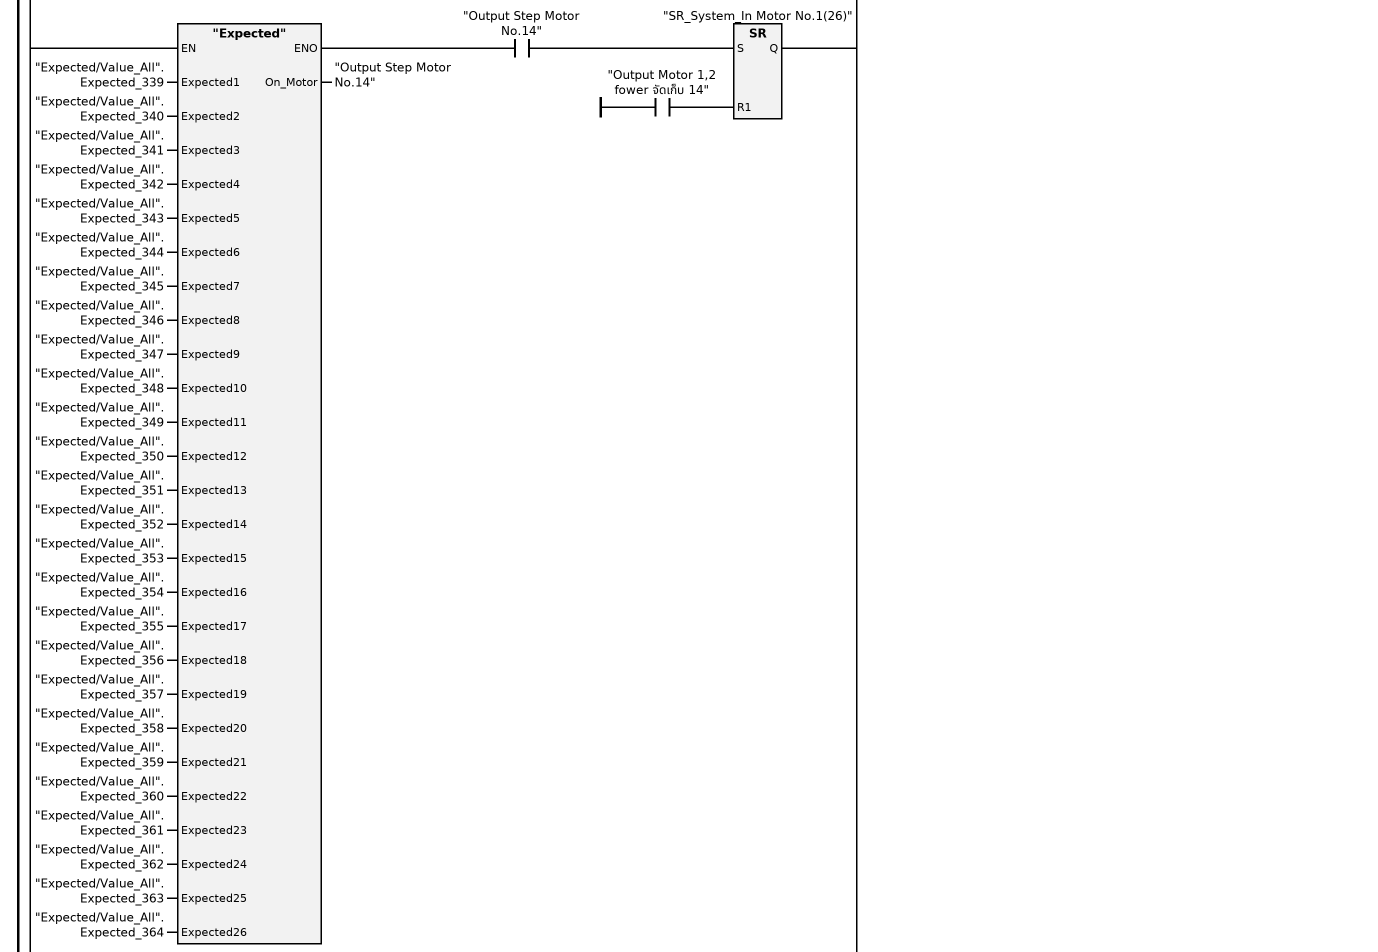
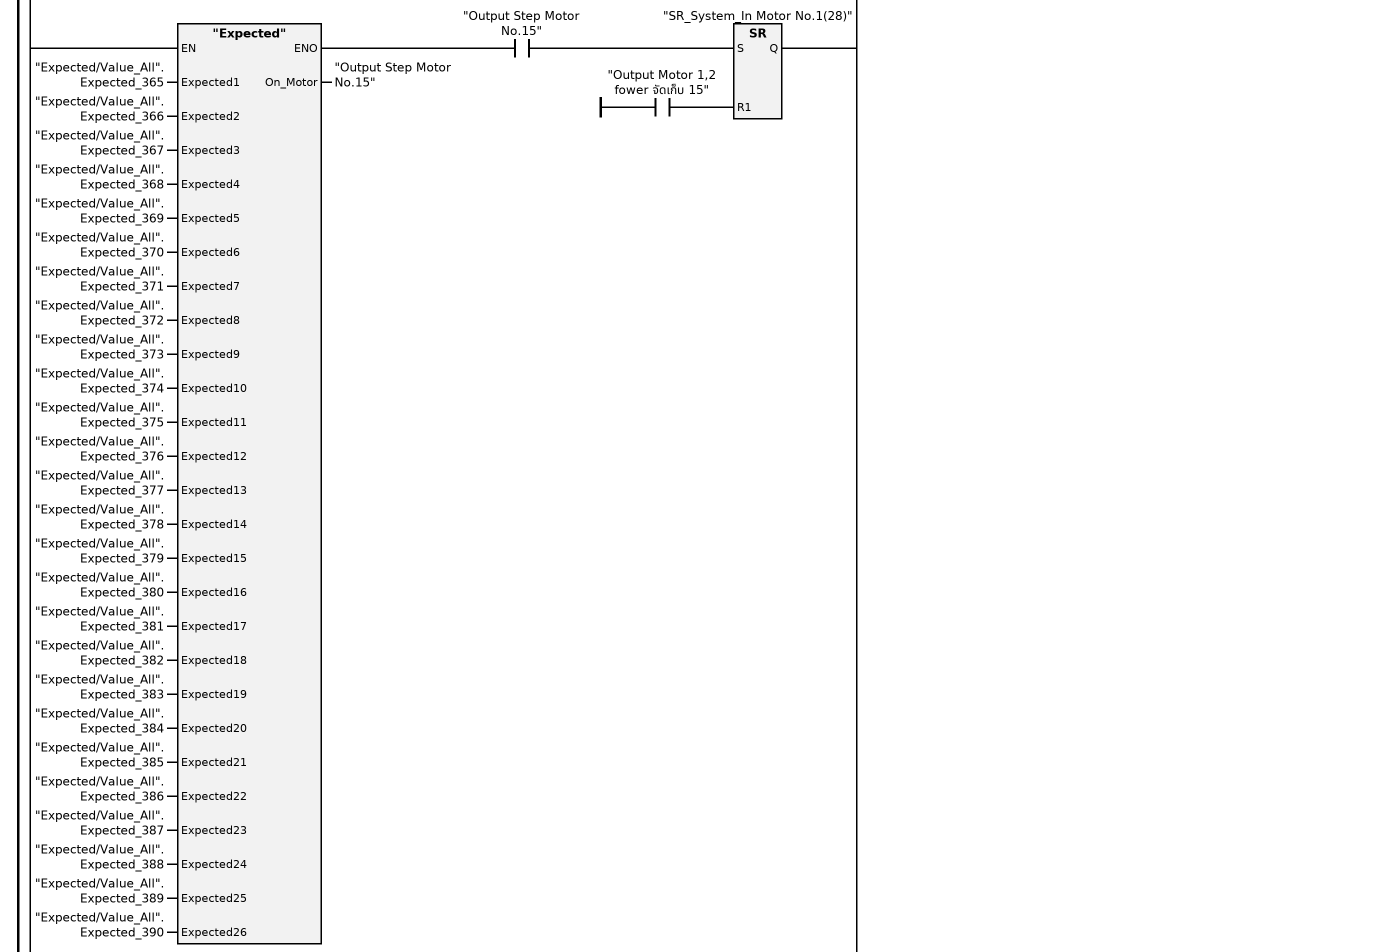
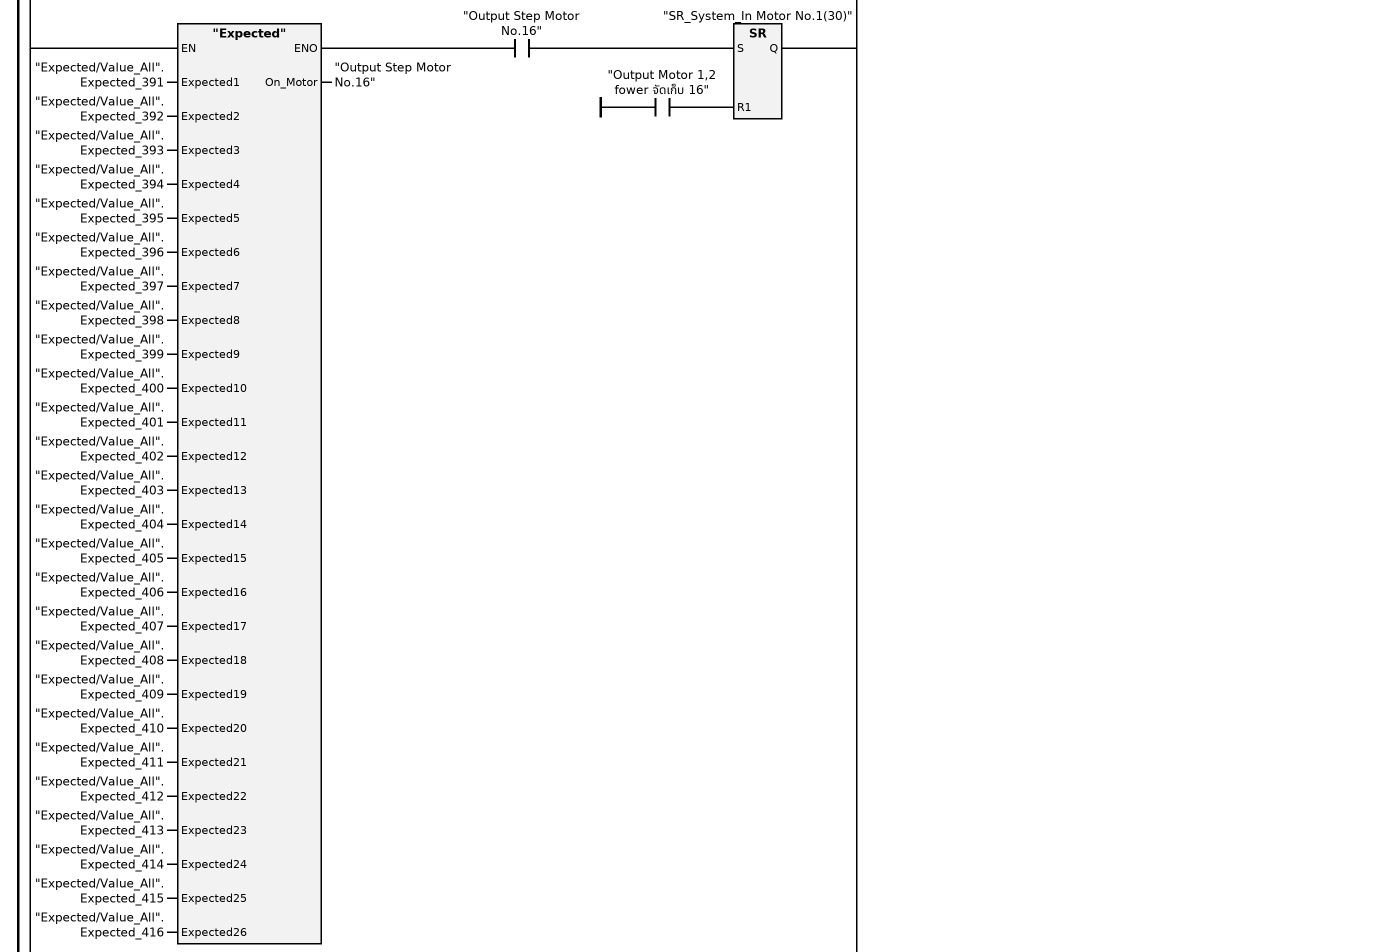
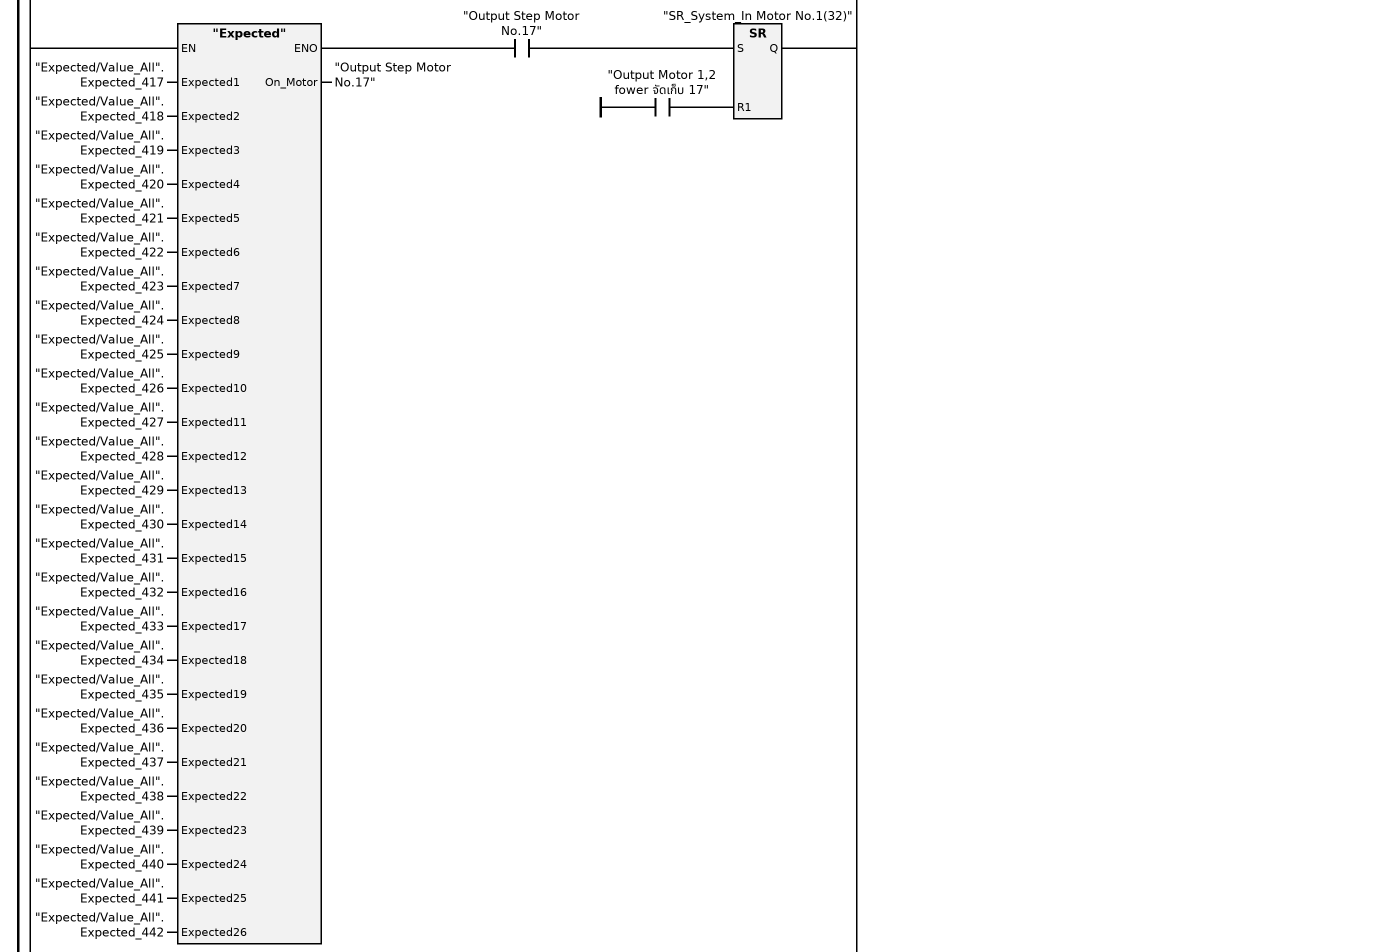
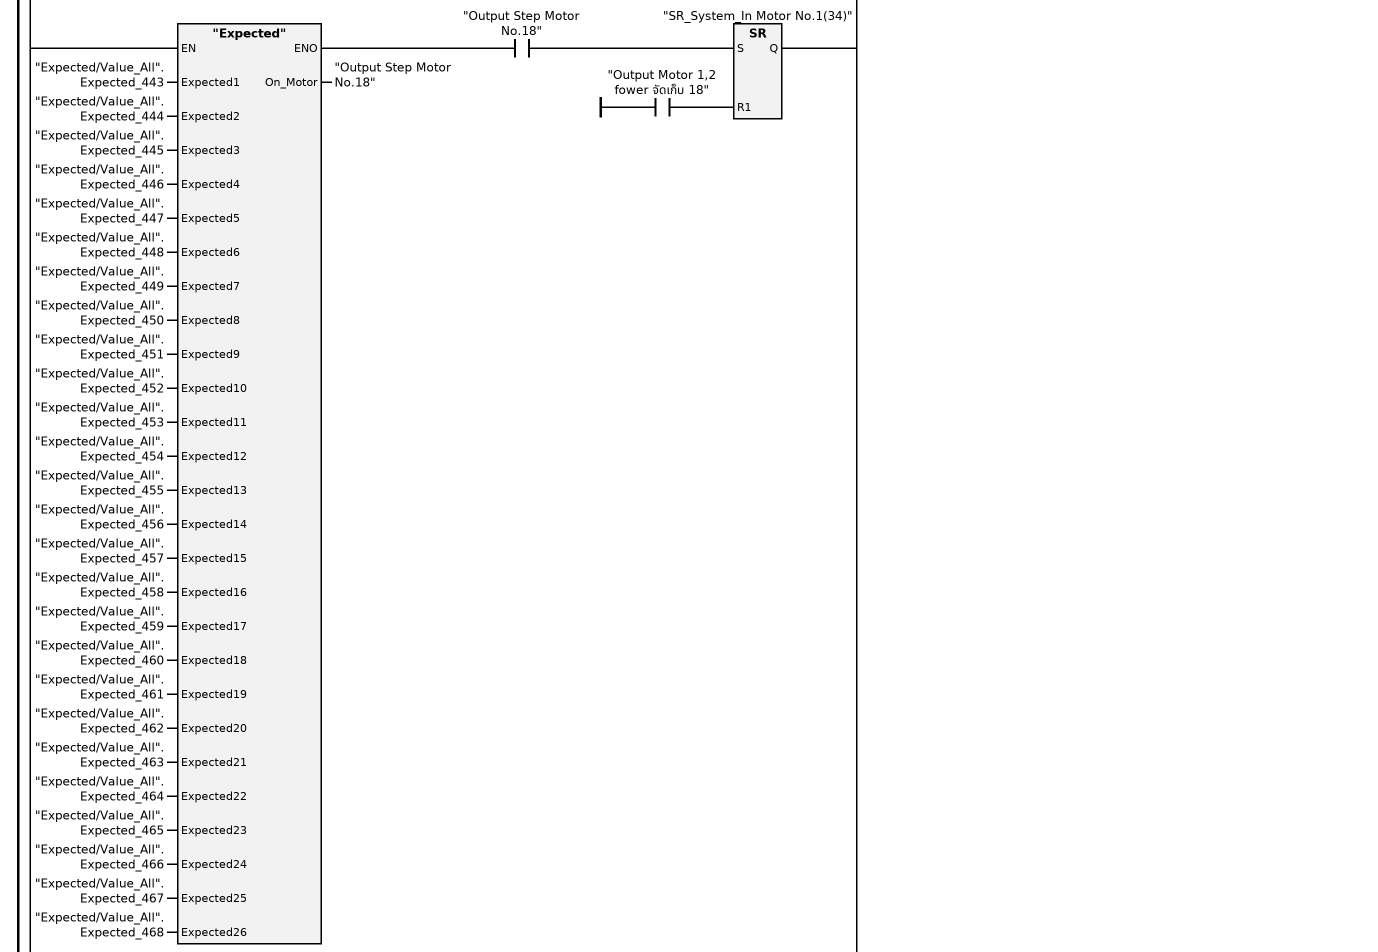
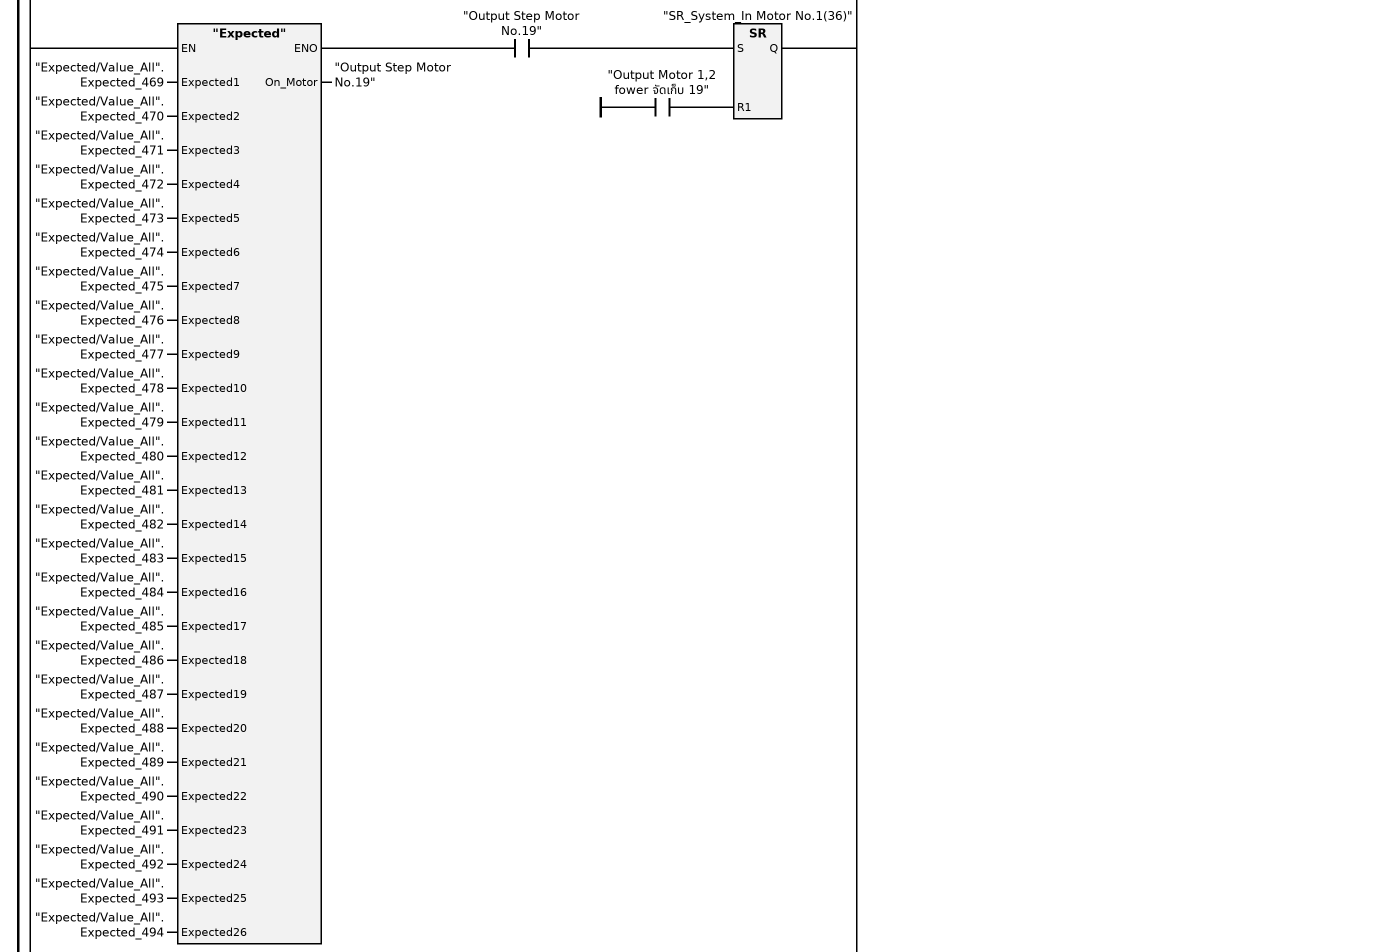
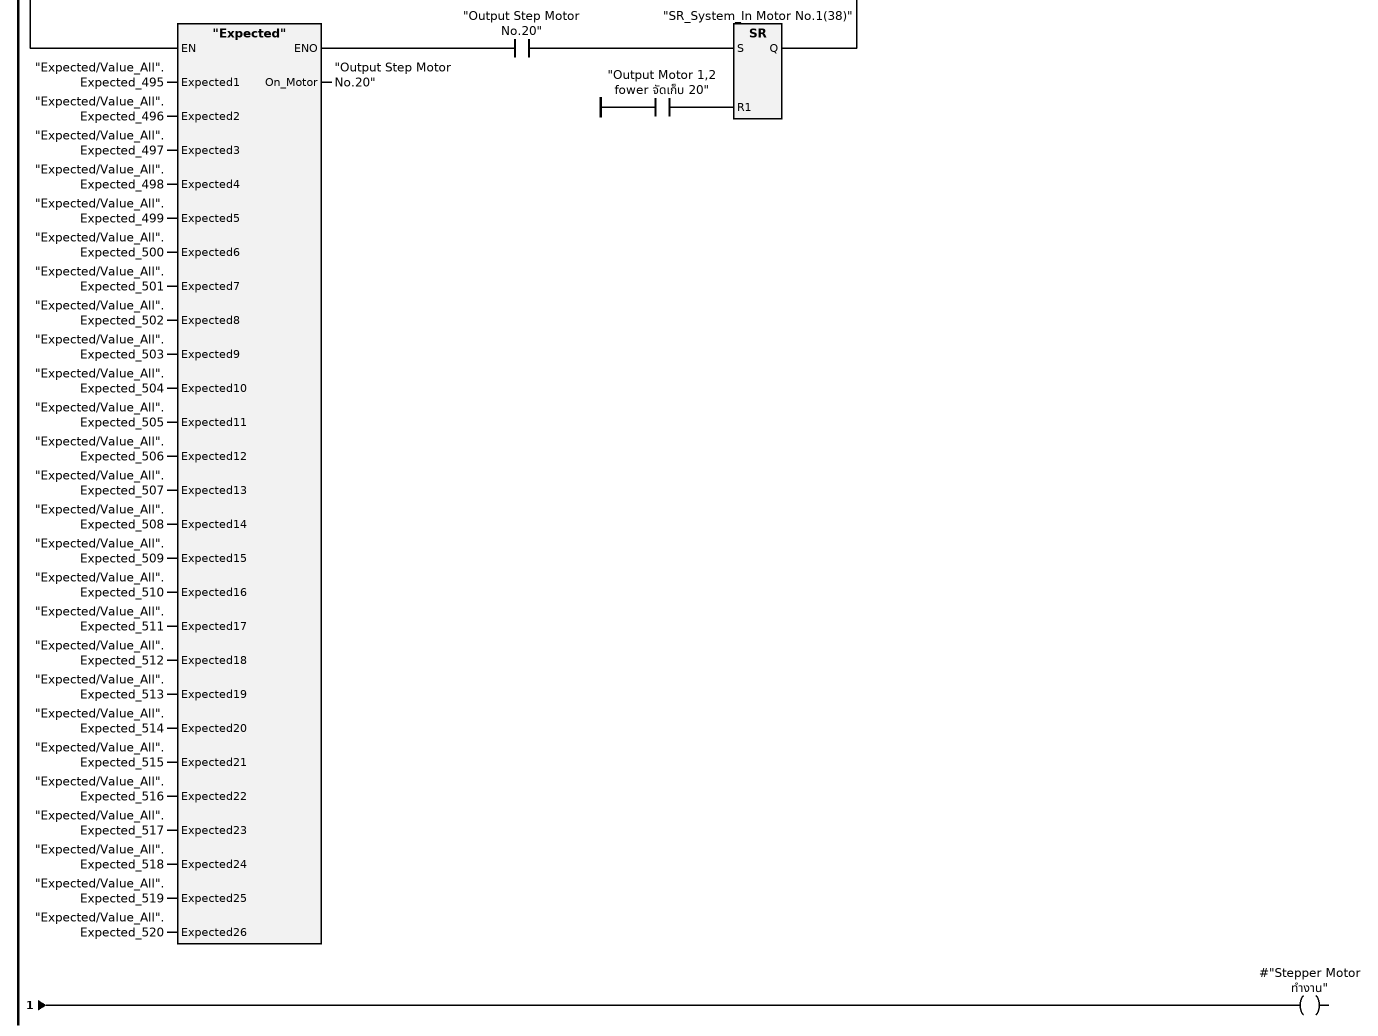
   RUNG wire#powerrail
      "Expected"(Expected1 := "Expected/Value_All".Expected_1, Expected2 := "Expected/Value_All".Expected_2, Expected3 := "Expected/Value_All".Expected_3, Expected4 := "Expected/Value_All".Expected_4, Expected5 := "Expected/Value_All".Expected_5, Expected6 := "Expected/Value_All".Expected_6, Expected7 := "Expected/Value_All".Expected_7, Expected8 := "Expected/Value_All".Expected_8, Expected9 := "Expected/Value_All".Expected_9, Expected10 := "Expected/Value_All".Expected_10, Expected11 := "Expected/Value_All".Expected_11, Expected12 := "Expected/Value_All".Expected_12, Expected13 := "Expected/Value_All".Expected_13, Expected14 := "Expected/Value_All".Expected_14, Expected15 := "Expected/Value_All".Expected_15, Expected16 := "Expected/Value_All".Expected_16, Expected17 := "Expected/Value_All".Expected_17, Expected18 := "Expected/Value_All".Expected_18, Expected19 := "Expected/Value_All".Expected_19, Expected20 := "Expected/Value_All".Expected_20, Expected21 := "Expected/Value_All".Expected_21, Expected22 := "Expected/Value_All".Expected_22, Expected23 := "Expected/Value_All".Expected_23, Expected24 := "Expected/Value_All".Expected_24, Expected25 := "Expected/Value_All".Expected_25, Expected26 := "Expected/Value_All".Expected_26, On_Motor => "Output Step Motor No.1")
      Contact( "Output Step Motor No.1" )
      S_SR(operand := "SR_System_In Motor No.1", r1 := wire#w1)
      wire#w2
      "test หลังเคลื่อนที่มาตำแหน่งปล่อยกล่องยา"()
      Contact( "หมุนไปตำแหต่งปล่อยกล่องยา" )
      Coil( #"Stepper Motor  ทำงาน" )
   END_RUNG
   RUNG wire#powerrail
      Contact( "Output Motor 1,2 fower จัดเก็บ 1" )
   END_RUNG wire#w1
   RUNG wire#powerrail
      "Expected"(Expected1 := "Expected/Value_All".Expected_27, Expected2 := "Expected/Value_All".Expected_28, Expected3 := "Expected/Value_All".Expected_29, Expected4 := "Expected/Value_All".Expected_30, Expected5 := "Expected/Value_All".Expected_31, Expected6 := "Expected/Value_All".Expected_32, Expected7 := "Expected/Value_All".Expected_33, Expected8 := "Expected/Value_All".Expected_34, Expected9 := "Expected/Value_All".Expected_35, Expected10 := "Expected/Value_All".Expected_36, Expected11 := "Expected/Value_All".Expected_37, Expected12 := "Expected/Value_All".Expected_38, Expected13 := "Expected/Value_All".Expected_39, Expected14 := "Expected/Value_All".Expected_40, Expected15 := "Expected/Value_All".Expected_41, Expected16 := "Expected/Value_All".Expected_42, Expected17 := "Expected/Value_All".Expected_43, Expected18 := "Expected/Value_All".Expected_44, Expected19 := "Expected/Value_All".Expected_45, Expected20 := "Expected/Value_All".Expected_46, Expected21 := "Expected/Value_All".Expected_47, Expected22 := "Expected/Value_All".Expected_48, Expected23 := "Expected/Value_All".Expected_49, Expected24 := "Expected/Value_All".Expected_50, Expected25 := "Expected/Value_All".Expected_51, Expected26 := "Expected/Value_All".Expected_52, On_Motor => "Output Step Motor No.2")
      Contact( "Output Step Motor No.2" )
      S_SR(operand := "SR_System_In Motor No.1(2)", r1 := wire#w3)
   END_RUNG wire#w2
   RUNG wire#powerrail
      Contact( "Output Motor 1,2 fower จัดเก็บ 2" )
   END_RUNG wire#w3
   RUNG wire#powerrail
      "Expected"(Expected1 := "Expected/Value_All".Expected_53, Expected2 := "Expected/Value_All".Expected_54, Expected3 := "Expected/Value_All".Expected_55, Expected4 := "Expected/Value_All".Expected_56, Expected5 := "Expected/Value_All".Expected_57, Expected6 := "Expected/Value_All".Expected_58, Expected7 := "Expected/Value_All".Expected_59, Expected8 := "Expected/Value_All".Expected_60, Expected9 := "Expected/Value_All".Expected_61, Expected10 := "Expected/Value_All".Expected_62, Expected11 := "Expected/Value_All".Expected_63, Expected12 := "Expected/Value_All".Expected_64, Expected13 := "Expected/Value_All".Expected_65, Expected14 := "Expected/Value_All".Expected_66, Expected15 := "Expected/Value_All".Expected_67, Expected16 := "Expected/Value_All".Expected_68, Expected17 := "Expected/Value_All".Expected_69, Expected18 := "Expected/Value_All".Expected_70, Expected19 := "Expected/Value_All".Expected_71, Expected20 := "Expected/Value_All".Expected_72, Expected21 := "Expected/Value_All".Expected_73, Expected22 := "Expected/Value_All".Expected_74, Expected23 := "Expected/Value_All".Expected_75, Expected24 := "Expected/Value_All".Expected_76, Expected25 := "Expected/Value_All".Expected_77, Expected26 := "Expected/Value_All".Expected_78, On_Motor => "Output Step Motor No.3")
      Contact( "Output Step Motor No.3" )
      S_SR(operand := "SR_System_In Motor No.1(4)", r1 := wire#w4)
   END_RUNG wire#w2
   RUNG wire#powerrail
      Contact( "Output Motor 1,2 fower จัดเก็บ 3" )
   END_RUNG wire#w4
   RUNG wire#powerrail
      "Expected"(Expected1 := "Expected/Value_All".Expected_79, Expected2 := "Expected/Value_All".Expected_80, Expected3 := "Expected/Value_All".Expected_81, Expected4 := "Expected/Value_All".Expected_82, Expected5 := "Expected/Value_All".Expected_83, Expected6 := "Expected/Value_All".Expected_84, Expected7 := "Expected/Value_All".Expected_85, Expected8 := "Expected/Value_All".Expected_86, Expected9 := "Expected/Value_All".Expected_87, Expected10 := "Expected/Value_All".Expected_88, Expected11 := "Expected/Value_All".Expected_89, Expected12 := "Expected/Value_All".Expected_90, Expected13 := "Expected/Value_All".Expected_91, Expected14 := "Expected/Value_All".Expected_92, Expected15 := "Expected/Value_All".Expected_93, Expected16 := "Expected/Value_All".Expected_94, Expected17 := "Expected/Value_All".Expected_95, Expected18 := "Expected/Value_All".Expected_96, Expected19 := "Expected/Value_All".Expected_97, Expected20 := "Expected/Value_All".Expected_98, Expected21 := "Expected/Value_All".Expected_99, Expected22 := "Expected/Value_All".Expected_100, Expected23 := "Expected/Value_All".Expected_101, Expected24 := "Expected/Value_All".Expected_102, Expected25 := "Expected/Value_All".Expected_103, Expected26 := "Expected/Value_All".Expected_104, On_Motor => "Output Step Motor No.4")
      Contact( "Output Step Motor No.4" )
      S_SR(operand := "SR_System_In Motor No.1(6)", r1 := wire#w5)
   END_RUNG wire#w2
   RUNG wire#powerrail
      Contact( "Output Motor 1,2 fower จัดเก็บ 4" )
   END_RUNG wire#w5
   RUNG wire#powerrail
      "Expected"(Expected1 := "Expected/Value_All".Expected_105, Expected2 := "Expected/Value_All".Expected_106, Expected3 := "Expected/Value_All".Expected_107, Expected4 := "Expected/Value_All".Expected_108, Expected5 := "Expected/Value_All".Expected_109, Expected6 := "Expected/Value_All".Expected_110, Expected7 := "Expected/Value_All".Expected_111, Expected8 := "Expected/Value_All".Expected_112, Expected9 := "Expected/Value_All".Expected_113, Expected10 := "Expected/Value_All".Expected_114, Expected11 := "Expected/Value_All".Expected_115, Expected12 := "Expected/Value_All".Expected_116, Expected13 := "Expected/Value_All".Expected_117, Expected14 := "Expected/Value_All".Expected_118, Expected15 := "Expected/Value_All".Expected_119, Expected16 := "Expected/Value_All".Expected_120, Expected17 := "Expected/Value_All".Expected_121, Expected18 := "Expected/Value_All".Expected_122, Expected19 := "Expected/Value_All".Expected_123, Expected20 := "Expected/Value_All".Expected_124, Expected21 := "Expected/Value_All".Expected_125, Expected22 := "Expected/Value_All".Expected_126, Expected23 := "Expected/Value_All".Expected_127, Expected24 := "Expected/Value_All".Expected_128, Expected25 := "Expected/Value_All".Expected_129, Expected26 := "Expected/Value_All".Expected_130, On_Motor => "Output Step Motor No.5")
      Contact( "Output Step Motor No.5" )
      S_SR(operand := "SR_System_In Motor No.1(8)", r1 := wire#w6)
   END_RUNG wire#w2
   RUNG wire#powerrail
      Contact( "Output Motor 1,2 fower จัดเก็บ 5" )
   END_RUNG wire#w6
   RUNG wire#powerrail
      "Expected"(Expected1 := "Expected/Value_All".Expected_131, Expected2 := "Expected/Value_All".Expected_132, Expected3 := "Expected/Value_All".Expected_133, Expected4 := "Expected/Value_All".Expected_134, Expected5 := "Expected/Value_All".Expected_135, Expected6 := "Expected/Value_All".Expected_136, Expected7 := "Expected/Value_All".Expected_137, Expected8 := "Expected/Value_All".Expected_138, Expected9 := "Expected/Value_All".Expected_139, Expected10 := "Expected/Value_All".Expected_140, Expected11 := "Expected/Value_All".Expected_141, Expected12 := "Expected/Value_All".Expected_142, Expected13 := "Expected/Value_All".Expected_143, Expected14 := "Expected/Value_All".Expected_144, Expected15 := "Expected/Value_All".Expected_145, Expected16 := "Expected/Value_All".Expected_146, Expected17 := "Expected/Value_All".Expected_147, Expected18 := "Expected/Value_All".Expected_148, Expected19 := "Expected/Value_All".Expected_149, Expected20 := "Expected/Value_All".Expected_150, Expected21 := "Expected/Value_All".Expected_151, Expected22 := "Expected/Value_All".Expected_152, Expected23 := "Expected/Value_All".Expected_153, Expected24 := "Expected/Value_All".Expected_154, Expected25 := "Expected/Value_All".Expected_155, Expected26 := "Expected/Value_All".Expected_156, On_Motor => "Output Step Motor No.6")
      Contact( "Output Step Motor No.6" )
      S_SR(operand := "SR_System_In Motor No.1(10)", r1 := wire#w7)
   END_RUNG wire#w2
   RUNG wire#powerrail
      Contact( "Output Motor 1,2 fower จัดเก็บ 6" )
   END_RUNG wire#w7
   RUNG wire#powerrail
      "Expected"(Expected1 := "Expected/Value_All".Expected_157, Expected2 := "Expected/Value_All".Expected_158, Expected3 := "Expected/Value_All".Expected_159, Expected4 := "Expected/Value_All".Expected_160, Expected5 := "Expected/Value_All".Expected_161, Expected6 := "Expected/Value_All".Expected_162, Expected7 := "Expected/Value_All".Expected_163, Expected8 := "Expected/Value_All".Expected_164, Expected9 := "Expected/Value_All".Expected_165, Expected10 := "Expected/Value_All".Expected_166, Expected11 := "Expected/Value_All".Expected_167, Expected12 := "Expected/Value_All".Expected_168, Expected13 := "Expected/Value_All".Expected_169, Expected14 := "Expected/Value_All".Expected_170, Expected15 := "Expected/Value_All".Expected_171, Expected16 := "Expected/Value_All".Expected_172, Expected17 := "Expected/Value_All".Expected_173, Expected18 := "Expected/Value_All".Expected_174, Expected19 := "Expected/Value_All".Expected_175, Expected20 := "Expected/Value_All".Expected_176, Expected21 := "Expected/Value_All".Expected_177, Expected22 := "Expected/Value_All".Expected_178, Expected23 := "Expected/Value_All".Expected_179, Expected24 := "Expected/Value_All".Expected_180, Expected25 := "Expected/Value_All".Expected_181, Expected26 := "Expected/Value_All".Expected_182, On_Motor => "Output Step Motor No.7")
      Contact( "Output Step Motor No.7" )
      S_SR(operand := "SR_System_In Motor No.1(12)", r1 := wire#w8)
   END_RUNG wire#w2
   RUNG wire#powerrail
      Contact( "Output Motor 1,2 fower จัดเก็บ 7" )
   END_RUNG wire#w8
   RUNG wire#powerrail
      "Expected"(Expected1 := "Expected/Value_All".Expected_183, Expected2 := "Expected/Value_All".Expected_184, Expected3 := "Expected/Value_All".Expected_185, Expected4 := "Expected/Value_All".Expected_186, Expected5 := "Expected/Value_All".Expected_187, Expected6 := "Expected/Value_All".Expected_188, Expected7 := "Expected/Value_All".Expected_189, Expected8 := "Expected/Value_All".Expected_190, Expected9 := "Expected/Value_All".Expected_191, Expected10 := "Expected/Value_All".Expected_192, Expected11 := "Expected/Value_All".Expected_193, Expected12 := "Expected/Value_All".Expected_194, Expected13 := "Expected/Value_All".Expected_195, Expected14 := "Expected/Value_All".Expected_196, Expected15 := "Expected/Value_All".Expected_197, Expected16 := "Expected/Value_All".Expected_198, Expected17 := "Expected/Value_All".Expected_199, Expected18 := "Expected/Value_All".Expected_200, Expected19 := "Expected/Value_All".Expected_201, Expected20 := "Expected/Value_All".Expected_202, Expected21 := "Expected/Value_All".Expected_203, Expected22 := "Expected/Value_All".Expected_204, Expected23 := "Expected/Value_All".Expected_205, Expected24 := "Expected/Value_All".Expected_206, Expected25 := "Expected/Value_All".Expected_207, Expected26 := "Expected/Value_All".Expected_208, On_Motor => "Output Step Motor No.8")
      Contact( "Output Step Motor No.8" )
      S_SR(operand := "SR_System_In Motor No.1(14)", r1 := wire#w9)
   END_RUNG wire#w2
   RUNG wire#powerrail
      Contact( "Output Motor 1,2 fower จัดเก็บ 8" )
   END_RUNG wire#w9
   RUNG wire#powerrail
      "Expected"(Expected1 := "Expected/Value_All".Expected_209, Expected2 := "Expected/Value_All".Expected_210, Expected3 := "Expected/Value_All".Expected_211, Expected4 := "Expected/Value_All".Expected_212, Expected5 := "Expected/Value_All".Expected_213, Expected6 := "Expected/Value_All".Expected_214, Expected7 := "Expected/Value_All".Expected_215, Expected8 := "Expected/Value_All".Expected_216, Expected9 := "Expected/Value_All".Expected_217, Expected10 := "Expected/Value_All".Expected_218, Expected11 := "Expected/Value_All".Expected_219, Expected12 := "Expected/Value_All".Expected_220, Expected13 := "Expected/Value_All".Expected_221, Expected14 := "Expected/Value_All".Expected_222, Expected15 := "Expected/Value_All".Expected_223, Expected16 := "Expected/Value_All".Expected_224, Expected17 := "Expected/Value_All".Expected_225, Expected18 := "Expected/Value_All".Expected_226, Expected19 := "Expected/Value_All".Expected_227, Expected20 := "Expected/Value_All".Expected_228, Expected21 := "Expected/Value_All".Expected_229, Expected22 := "Expected/Value_All".Expected_230, Expected23 := "Expected/Value_All".Expected_231, Expected24 := "Expected/Value_All".Expected_232, Expected25 := "Expected/Value_All".Expected_233, Expected26 := "Expected/Value_All".Expected_234, On_Motor => "Output Step Motor No.9")
      Contact( "Output Step Motor No.9" )
      S_SR(operand := "SR_System_In Motor No.1(16)", r1 := wire#w10)
   END_RUNG wire#w2
   RUNG wire#powerrail
      Contact( "Output Motor 1,2 fower จัดเก็บ 9" )
   END_RUNG wire#w10
   RUNG wire#powerrail
      "Expected"(Expected1 := "Expected/Value_All".Expected_235, Expected2 := "Expected/Value_All".Expected_236, Expected3 := "Expected/Value_All".Expected_237, Expected4 := "Expected/Value_All".Expected_238, Expected5 := "Expected/Value_All".Expected_239, Expected6 := "Expected/Value_All".Expected_240, Expected7 := "Expected/Value_All".Expected_241, Expected8 := "Expected/Value_All".Expected_242, Expected9 := "Expected/Value_All".Expected_243, Expected10 := "Expected/Value_All".Expected_244, Expected11 := "Expected/Value_All".Expected_245, Expected12 := "Expected/Value_All".Expected_246, Expected13 := "Expected/Value_All".Expected_247, Expected14 := "Expected/Value_All".Expected_248, Expected15 := "Expected/Value_All".Expected_249, Expected16 := "Expected/Value_All".Expected_250, Expected17 := "Expected/Value_All".Expected_251, Expected18 := "Expected/Value_All".Expected_252, Expected19 := "Expected/Value_All".Expected_253, Expected20 := "Expected/Value_All".Expected_254, Expected21 := "Expected/Value_All".Expected_255, Expected22 := "Expected/Value_All".Expected_256, Expected23 := "Expected/Value_All".Expected_257, Expected24 := "Expected/Value_All".Expected_258, Expected25 := "Expected/Value_All".Expected_259, Expected26 := "Expected/Value_All".Expected_260, On_Motor => "Output Step Motor No.10")
      Contact( "Output Step Motor No.10" )
      S_SR(operand := "SR_System_In Motor No.1(18)", r1 := wire#w11)
   END_RUNG wire#w2
   RUNG wire#powerrail
      Contact( "Output Motor 1,2 fower จัดเก็บ 10" )
   END_RUNG wire#w11
   RUNG wire#powerrail
      "Expected"(Expected1 := "Expected/Value_All".Expected_261, Expected2 := "Expected/Value_All".Expected_262, Expected3 := "Expected/Value_All".Expected_263, Expected4 := "Expected/Value_All".Expected_264, Expected5 := "Expected/Value_All".Expected_265, Expected6 := "Expected/Value_All".Expected_266, Expected7 := "Expected/Value_All".Expected_267, Expected8 := "Expected/Value_All".Expected_268, Expected9 := "Expected/Value_All".Expected_269, Expected10 := "Expected/Value_All".Expected_270, Expected11 := "Expected/Value_All".Expected_271, Expected12 := "Expected/Value_All".Expected_272, Expected13 := "Expected/Value_All".Expected_273, Expected14 := "Expected/Value_All".Expected_274, Expected15 := "Expected/Value_All".Expected_275, Expected16 := "Expected/Value_All".Expected_276, Expected17 := "Expected/Value_All".Expected_277, Expected18 := "Expected/Value_All".Expected_278, Expected19 := "Expected/Value_All".Expected_279, Expected20 := "Expected/Value_All".Expected_280, Expected21 := "Expected/Value_All".Expected_281, Expected22 := "Expected/Value_All".Expected_282, Expected23 := "Expected/Value_All".Expected_283, Expected24 := "Expected/Value_All".Expected_284, Expected25 := "Expected/Value_All".Expected_285, Expected26 := "Expected/Value_All".Expected_286, On_Motor => "Output Step Motor No.11")
      Contact( "Output Step Motor No.11" )
      S_SR(operand := "SR_System_In Motor No.1(20)", r1 := wire#w12)
   END_RUNG wire#w2
   RUNG wire#powerrail
      Contact( "Output Motor 1,2 fower จัดเก็บ 11" )
   END_RUNG wire#w12
   RUNG wire#powerrail
      "Expected"(Expected1 := "Expected/Value_All".Expected_287, Expected2 := "Expected/Value_All".Expected_288, Expected3 := "Expected/Value_All".Expected_289, Expected4 := "Expected/Value_All".Expected_290, Expected5 := "Expected/Value_All".Expected_291, Expected6 := "Expected/Value_All".Expected_292, Expected7 := "Expected/Value_All".Expected_293, Expected8 := "Expected/Value_All".Expected_294, Expected9 := "Expected/Value_All".Expected_295, Expected10 := "Expected/Value_All".Expected_296, Expected11 := "Expected/Value_All".Expected_297, Expected12 := "Expected/Value_All".Expected_298, Expected13 := "Expected/Value_All".Expected_299, Expected14 := "Expected/Value_All".Expected_300, Expected15 := "Expected/Value_All".Expected_301, Expected16 := "Expected/Value_All".Expected_302, Expected17 := "Expected/Value_All".Expected_303, Expected18 := "Expected/Value_All".Expected_304, Expected19 := "Expected/Value_All".Expected_305, Expected20 := "Expected/Value_All".Expected_306, Expected21 := "Expected/Value_All".Expected_307, Expected22 := "Expected/Value_All".Expected_308, Expected23 := "Expected/Value_All".Expected_309, Expected24 := "Expected/Value_All".Expected_310, Expected25 := "Expected/Value_All".Expected_311, Expected26 := "Expected/Value_All".Expected_312, On_Motor => "Output Step Motor No.12")
      Contact( "Output Step Motor No.12" )
      S_SR(operand := "SR_System_In Motor No.1(22)", r1 := wire#w13)
   END_RUNG wire#w2
   RUNG wire#powerrail
      Contact( "Output Motor 1,2 fower จัดเก็บ 12" )
   END_RUNG wire#w13
   RUNG wire#powerrail
      "Expected"(Expected1 := "Expected/Value_All".Expected_313, Expected2 := "Expected/Value_All".Expected_314, Expected3 := "Expected/Value_All".Expected_315, Expected4 := "Expected/Value_All".Expected_316, Expected5 := "Expected/Value_All".Expected_317, Expected6 := "Expected/Value_All".Expected_318, Expected7 := "Expected/Value_All".Expected_319, Expected8 := "Expected/Value_All".Expected_320, Expected9 := "Expected/Value_All".Expected_321, Expected10 := "Expected/Value_All".Expected_322, Expected11 := "Expected/Value_All".Expected_323, Expected12 := "Expected/Value_All".Expected_324, Expected13 := "Expected/Value_All".Expected_325, Expected14 := "Expected/Value_All".Expected_326, Expected15 := "Expected/Value_All".Expected_327, Expected16 := "Expected/Value_All".Expected_328, Expected17 := "Expected/Value_All".Expected_329, Expected18 := "Expected/Value_All".Expected_330, Expected19 := "Expected/Value_All".Expected_331, Expected20 := "Expected/Value_All".Expected_332, Expected21 := "Expected/Value_All".Expected_333, Expected22 := "Expected/Value_All".Expected_334, Expected23 := "Expected/Value_All".Expected_335, Expected24 := "Expected/Value_All".Expected_336, Expected25 := "Expected/Value_All".Expected_337, Expected26 := "Expected/Value_All".Expected_338, On_Motor => "Output Step Motor No.13")
      Contact( "Output Step Motor No.13" )
      S_SR(operand := "SR_System_In Motor No.1(24)", r1 := wire#w14)
   END_RUNG wire#w2
   RUNG wire#powerrail
      Contact( "Output Motor 1,2 fower จัดเก็บ 13" )
   END_RUNG wire#w14
   RUNG wire#powerrail
      "Expected"(Expected1 := "Expected/Value_All".Expected_339, Expected2 := "Expected/Value_All".Expected_340, Expected3 := "Expected/Value_All".Expected_341, Expected4 := "Expected/Value_All".Expected_342, Expected5 := "Expected/Value_All".Expected_343, Expected6 := "Expected/Value_All".Expected_344, Expected7 := "Expected/Value_All".Expected_345, Expected8 := "Expected/Value_All".Expected_346, Expected9 := "Expected/Value_All".Expected_347, Expected10 := "Expected/Value_All".Expected_348, Expected11 := "Expected/Value_All".Expected_349, Expected12 := "Expected/Value_All".Expected_350, Expected13 := "Expected/Value_All".Expected_351, Expected14 := "Expected/Value_All".Expected_352, Expected15 := "Expected/Value_All".Expected_353, Expected16 := "Expected/Value_All".Expected_354, Expected17 := "Expected/Value_All".Expected_355, Expected18 := "Expected/Value_All".Expected_356, Expected19 := "Expected/Value_All".Expected_357, Expected20 := "Expected/Value_All".Expected_358, Expected21 := "Expected/Value_All".Expected_359, Expected22 := "Expected/Value_All".Expected_360, Expected23 := "Expected/Value_All".Expected_361, Expected24 := "Expected/Value_All".Expected_362, Expected25 := "Expected/Value_All".Expected_363, Expected26 := "Expected/Value_All".Expected_364, On_Motor => "Output Step Motor No.14")
      Contact( "Output Step Motor No.14" )
      S_SR(operand := "SR_System_In Motor No.1(26)", r1 := wire#w15)
   END_RUNG wire#w2
   RUNG wire#powerrail
      Contact( "Output Motor 1,2 fower จัดเก็บ 14" )
   END_RUNG wire#w15
   RUNG wire#powerrail
      "Expected"(Expected1 := "Expected/Value_All".Expected_365, Expected2 := "Expected/Value_All".Expected_366, Expected3 := "Expected/Value_All".Expected_367, Expected4 := "Expected/Value_All".Expected_368, Expected5 := "Expected/Value_All".Expected_369, Expected6 := "Expected/Value_All".Expected_370, Expected7 := "Expected/Value_All".Expected_371, Expected8 := "Expected/Value_All".Expected_372, Expected9 := "Expected/Value_All".Expected_373, Expected10 := "Expected/Value_All".Expected_374, Expected11 := "Expected/Value_All".Expected_375, Expected12 := "Expected/Value_All".Expected_376, Expected13 := "Expected/Value_All".Expected_377, Expected14 := "Expected/Value_All".Expected_378, Expected15 := "Expected/Value_All".Expected_379, Expected16 := "Expected/Value_All".Expected_380, Expected17 := "Expected/Value_All".Expected_381, Expected18 := "Expected/Value_All".Expected_382, Expected19 := "Expected/Value_All".Expected_383, Expected20 := "Expected/Value_All".Expected_384, Expected21 := "Expected/Value_All".Expected_385, Expected22 := "Expected/Value_All".Expected_386, Expected23 := "Expected/Value_All".Expected_387, Expected24 := "Expected/Value_All".Expected_388, Expected25 := "Expected/Value_All".Expected_389, Expected26 := "Expected/Value_All".Expected_390, On_Motor => "Output Step Motor No.15")
      Contact( "Output Step Motor No.15" )
      S_SR(operand := "SR_System_In Motor No.1(28)", r1 := wire#w16)
   END_RUNG wire#w2
   RUNG wire#powerrail
      Contact( "Output Motor 1,2 fower จัดเก็บ 15" )
   END_RUNG wire#w16
   RUNG wire#powerrail
      "Expected"(Expected1 := "Expected/Value_All".Expected_391, Expected2 := "Expected/Value_All".Expected_392, Expected3 := "Expected/Value_All".Expected_393, Expected4 := "Expected/Value_All".Expected_394, Expected5 := "Expected/Value_All".Expected_395, Expected6 := "Expected/Value_All".Expected_396, Expected7 := "Expected/Value_All".Expected_397, Expected8 := "Expected/Value_All".Expected_398, Expected9 := "Expected/Value_All".Expected_399, Expected10 := "Expected/Value_All".Expected_400, Expected11 := "Expected/Value_All".Expected_401, Expected12 := "Expected/Value_All".Expected_402, Expected13 := "Expected/Value_All".Expected_403, Expected14 := "Expected/Value_All".Expected_404, Expected15 := "Expected/Value_All".Expected_405, Expected16 := "Expected/Value_All".Expected_406, Expected17 := "Expected/Value_All".Expected_407, Expected18 := "Expected/Value_All".Expected_408, Expected19 := "Expected/Value_All".Expected_409, Expected20 := "Expected/Value_All".Expected_410, Expected21 := "Expected/Value_All".Expected_411, Expected22 := "Expected/Value_All".Expected_412, Expected23 := "Expected/Value_All".Expected_413, Expected24 := "Expected/Value_All".Expected_414, Expected25 := "Expected/Value_All".Expected_415, Expected26 := "Expected/Value_All".Expected_416, On_Motor => "Output Step Motor No.16")
      Contact( "Output Step Motor No.16" )
      S_SR(operand := "SR_System_In Motor No.1(30)", r1 := wire#w17)
   END_RUNG wire#w2
   RUNG wire#powerrail
      Contact( "Output Motor 1,2 fower จัดเก็บ 16" )
   END_RUNG wire#w17
   RUNG wire#powerrail
      "Expected"(Expected1 := "Expected/Value_All".Expected_417, Expected2 := "Expected/Value_All".Expected_418, Expected3 := "Expected/Value_All".Expected_419, Expected4 := "Expected/Value_All".Expected_420, Expected5 := "Expected/Value_All".Expected_421, Expected6 := "Expected/Value_All".Expected_422, Expected7 := "Expected/Value_All".Expected_423, Expected8 := "Expected/Value_All".Expected_424, Expected9 := "Expected/Value_All".Expected_425, Expected10 := "Expected/Value_All".Expected_426, Expected11 := "Expected/Value_All".Expected_427, Expected12 := "Expected/Value_All".Expected_428, Expected13 := "Expected/Value_All".Expected_429, Expected14 := "Expected/Value_All".Expected_430, Expected15 := "Expected/Value_All".Expected_431, Expected16 := "Expected/Value_All".Expected_432, Expected17 := "Expected/Value_All".Expected_433, Expected18 := "Expected/Value_All".Expected_434, Expected19 := "Expected/Value_All".Expected_435, Expected20 := "Expected/Value_All".Expected_436, Expected21 := "Expected/Value_All".Expected_437, Expected22 := "Expected/Value_All".Expected_438, Expected23 := "Expected/Value_All".Expected_439, Expected24 := "Expected/Value_All".Expected_440, Expected25 := "Expected/Value_All".Expected_441, Expected26 := "Expected/Value_All".Expected_442, On_Motor => "Output Step Motor No.17")
      Contact( "Output Step Motor No.17" )
      S_SR(operand := "SR_System_In Motor No.1(32)", r1 := wire#w18)
   END_RUNG wire#w2
   RUNG wire#powerrail
      Contact( "Output Motor 1,2 fower จัดเก็บ 17" )
   END_RUNG wire#w18
   RUNG wire#powerrail
      "Expected"(Expected1 := "Expected/Value_All".Expected_443, Expected2 := "Expected/Value_All".Expected_444, Expected3 := "Expected/Value_All".Expected_445, Expected4 := "Expected/Value_All".Expected_446, Expected5 := "Expected/Value_All".Expected_447, Expected6 := "Expected/Value_All".Expected_448, Expected7 := "Expected/Value_All".Expected_449, Expected8 := "Expected/Value_All".Expected_450, Expected9 := "Expected/Value_All".Expected_451, Expected10 := "Expected/Value_All".Expected_452, Expected11 := "Expected/Value_All".Expected_453, Expected12 := "Expected/Value_All".Expected_454, Expected13 := "Expected/Value_All".Expected_455, Expected14 := "Expected/Value_All".Expected_456, Expected15 := "Expected/Value_All".Expected_457, Expected16 := "Expected/Value_All".Expected_458, Expected17 := "Expected/Value_All".Expected_459, Expected18 := "Expected/Value_All".Expected_460, Expected19 := "Expected/Value_All".Expected_461, Expected20 := "Expected/Value_All".Expected_462, Expected21 := "Expected/Value_All".Expected_463, Expected22 := "Expected/Value_All".Expected_464, Expected23 := "Expected/Value_All".Expected_465, Expected24 := "Expected/Value_All".Expected_466, Expected25 := "Expected/Value_All".Expected_467, Expected26 := "Expected/Value_All".Expected_468, On_Motor => "Output Step Motor No.18")
      Contact( "Output Step Motor No.18" )
      S_SR(operand := "SR_System_In Motor No.1(34)", r1 := wire#w19)
   END_RUNG wire#w2
   RUNG wire#powerrail
      Contact( "Output Motor 1,2 fower จัดเก็บ 18" )
   END_RUNG wire#w19
   RUNG wire#powerrail
      "Expected"(Expected1 := "Expected/Value_All".Expected_469, Expected2 := "Expected/Value_All".Expected_470, Expected3 := "Expected/Value_All".Expected_471, Expected4 := "Expected/Value_All".Expected_472, Expected5 := "Expected/Value_All".Expected_473, Expected6 := "Expected/Value_All".Expected_474, Expected7 := "Expected/Value_All".Expected_475, Expected8 := "Expected/Value_All".Expected_476, Expected9 := "Expected/Value_All".Expected_477, Expected10 := "Expected/Value_All".Expected_478, Expected11 := "Expected/Value_All".Expected_479, Expected12 := "Expected/Value_All".Expected_480, Expected13 := "Expected/Value_All".Expected_481, Expected14 := "Expected/Value_All".Expected_482, Expected15 := "Expected/Value_All".Expected_483, Expected16 := "Expected/Value_All".Expected_484, Expected17 := "Expected/Value_All".Expected_485, Expected18 := "Expected/Value_All".Expected_486, Expected19 := "Expected/Value_All".Expected_487, Expected20 := "Expected/Value_All".Expected_488, Expected21 := "Expected/Value_All".Expected_489, Expected22 := "Expected/Value_All".Expected_490, Expected23 := "Expected/Value_All".Expected_491, Expected24 := "Expected/Value_All".Expected_492, Expected25 := "Expected/Value_All".Expected_493, Expected26 := "Expected/Value_All".Expected_494, On_Motor => "Output Step Motor No.19")
      Contact( "Output Step Motor No.19" )
      S_SR(operand := "SR_System_In Motor No.1(36)", r1 := wire#w20)
   END_RUNG wire#w2
   RUNG wire#powerrail
      Contact( "Output Motor 1,2 fower จัดเก็บ 19" )
   END_RUNG wire#w20
   RUNG wire#powerrail
      "Expected"(Expected1 := "Expected/Value_All".Expected_495, Expected2 := "Expected/Value_All".Expected_496, Expected3 := "Expected/Value_All".Expected_497, Expected4 := "Expected/Value_All".Expected_498, Expected5 := "Expected/Value_All".Expected_499, Expected6 := "Expected/Value_All".Expected_500, Expected7 := "Expected/Value_All".Expected_501, Expected8 := "Expected/Value_All".Expected_502, Expected9 := "Expected/Value_All".Expected_503, Expected10 := "Expected/Value_All".Expected_504, Expected11 := "Expected/Value_All".Expected_505, Expected12 := "Expected/Value_All".Expected_506, Expected13 := "Expected/Value_All".Expected_507, Expected14 := "Expected/Value_All".Expected_508, Expected15 := "Expected/Value_All".Expected_509, Expected16 := "Expected/Value_All".Expected_510, Expected17 := "Expected/Value_All".Expected_511, Expected18 := "Expected/Value_All".Expected_512, Expected19 := "Expected/Value_All".Expected_513, Expected20 := "Expected/Value_All".Expected_514, Expected21 := "Expected/Value_All".Expected_515, Expected22 := "Expected/Value_All".Expected_516, Expected23 := "Expected/Value_All".Expected_517, Expected24 := "Expected/Value_All".Expected_518, Expected25 := "Expected/Value_All".Expected_519, Expected26 := "Expected/Value_All".Expected_520, On_Motor => "Output Step Motor No.20")
      Contact( "Output Step Motor No.20" )
      S_SR(operand := "SR_System_In Motor No.1(38)", r1 := wire#w21)
   END_RUNG wire#w2
   RUNG wire#powerrail
      Contact( "Output Motor 1,2 fower จัดเก็บ 20" )
   END_RUNG wire#w21
   // the same network as SCL:
   "Expected"(Expected1 := "Expected/Value_All".Expected_1,
              Expected2 := "Expected/Value_All".Expected_2,
              Expected3 := "Expected/Value_All".Expected_3,
              Expected4 := "Expected/Value_All".Expected_4,
              Expected5 := "Expected/Value_All".Expected_5,
              Expected6 := "Expected/Value_All".Expected_6,
              Expected7 := "Expected/Value_All".Expected_7,
              Expected8 := "Expected/Value_All".Expected_8,
              Expected9 := "Expected/Value_All".Expected_9,
              Expected10 := "Expected/Value_All".Expected_10,
              Expected11 := "Expected/Value_All".Expected_11,
              Expected12 := "Expected/Value_All".Expected_12,
              Expected13 := "Expected/Value_All".Expected_13,
              Expected14 := "Expected/Value_All".Expected_14,
              Expected15 := "Expected/Value_All".Expected_15,
              Expected16 := "Expected/Value_All".Expected_16,
              Expected17 := "Expected/Value_All".Expected_17,
              Expected18 := "Expected/Value_All".Expected_18,
              Expected19 := "Expected/Value_All".Expected_19,
              Expected20 := "Expected/Value_All".Expected_20,
              Expected21 := "Expected/Value_All".Expected_21,
              Expected22 := "Expected/Value_All".Expected_22,
              Expected23 := "Expected/Value_All".Expected_23,
              Expected24 := "Expected/Value_All".Expected_24,
              Expected25 := "Expected/Value_All".Expected_25,
              Expected26 := "Expected/Value_All".Expected_26,
              On_Motor => "Output Step Motor No.1",
              ENO => #_w1);
   IF #_w1 AND "Output Step Motor No.1" THEN
       "SR_System_In Motor No.1" := TRUE;   // SR flip-flop
   END_IF;
   IF "Output Motor 1,2 fower จัดเก็บ 1" THEN "SR_System_In Motor No.1" := FALSE; END_IF;
   #_w3 := "SR_System_In Motor No.1";
   "Expected"(Expected1 := "Expected/Value_All".Expected_27,
              Expected2 := "Expected/Value_All".Expected_28,
              Expected3 := "Expected/Value_All".Expected_29,
              Expected4 := "Expected/Value_All".Expected_30,
              Expected5 := "Expected/Value_All".Expected_31,
              Expected6 := "Expected/Value_All".Expected_32,
              Expected7 := "Expected/Value_All".Expected_33,
              Expected8 := "Expected/Value_All".Expected_34,
              Expected9 := "Expected/Value_All".Expected_35,
              Expected10 := "Expected/Value_All".Expected_36,
              Expected11 := "Expected/Value_All".Expected_37,
              Expected12 := "Expected/Value_All".Expected_38,
              Expected13 := "Expected/Value_All".Expected_39,
              Expected14 := "Expected/Value_All".Expected_40,
              Expected15 := "Expected/Value_All".Expected_41,
              Expected16 := "Expected/Value_All".Expected_42,
              Expected17 := "Expected/Value_All".Expected_43,
              Expected18 := "Expected/Value_All".Expected_44,
              Expected19 := "Expected/Value_All".Expected_45,
              Expected20 := "Expected/Value_All".Expected_46,
              Expected21 := "Expected/Value_All".Expected_47,
              Expected22 := "Expected/Value_All".Expected_48,
              Expected23 := "Expected/Value_All".Expected_49,
              Expected24 := "Expected/Value_All".Expected_50,
              Expected25 := "Expected/Value_All".Expected_51,
              Expected26 := "Expected/Value_All".Expected_52,
              On_Motor => "Output Step Motor No.2",
              ENO => #_w2);
   IF #_w2 AND "Output Step Motor No.2" THEN
       "SR_System_In Motor No.1(2)" := TRUE;   // SR flip-flop
   END_IF;
   IF "Output Motor 1,2 fower จัดเก็บ 2" THEN "SR_System_In Motor No.1(2)" := FALSE; END_IF;
   #_w5 := "SR_System_In Motor No.1(2)";
   "Expected"(Expected1 := "Expected/Value_All".Expected_53,
              Expected2 := "Expected/Value_All".Expected_54,
              Expected3 := "Expected/Value_All".Expected_55,
              Expected4 := "Expected/Value_All".Expected_56,
              Expected5 := "Expected/Value_All".Expected_57,
              Expected6 := "Expected/Value_All".Expected_58,
              Expected7 := "Expected/Value_All".Expected_59,
              Expected8 := "Expected/Value_All".Expected_60,
              Expected9 := "Expected/Value_All".Expected_61,
              Expected10 := "Expected/Value_All".Expected_62,
              Expected11 := "Expected/Value_All".Expected_63,
              Expected12 := "Expected/Value_All".Expected_64,
              Expected13 := "Expected/Value_All".Expected_65,
              Expected14 := "Expected/Value_All".Expected_66,
              Expected15 := "Expected/Value_All".Expected_67,
              Expected16 := "Expected/Value_All".Expected_68,
              Expected17 := "Expected/Value_All".Expected_69,
              Expected18 := "Expected/Value_All".Expected_70,
              Expected19 := "Expected/Value_All".Expected_71,
              Expected20 := "Expected/Value_All".Expected_72,
              Expected21 := "Expected/Value_All".Expected_73,
              Expected22 := "Expected/Value_All".Expected_74,
              Expected23 := "Expected/Value_All".Expected_75,
              Expected24 := "Expected/Value_All".Expected_76,
              Expected25 := "Expected/Value_All".Expected_77,
              Expected26 := "Expected/Value_All".Expected_78,
              On_Motor => "Output Step Motor No.3",
              ENO => #_w4);
   IF #_w4 AND "Output Step Motor No.3" THEN
       "SR_System_In Motor No.1(4)" := TRUE;   // SR flip-flop
   END_IF;
   IF "Output Motor 1,2 fower จัดเก็บ 3" THEN "SR_System_In Motor No.1(4)" := FALSE; END_IF;
   #_w7 := "SR_System_In Motor No.1(4)";
   "Expected"(Expected1 := "Expected/Value_All".Expected_79,
              Expected2 := "Expected/Value_All".Expected_80,
              Expected3 := "Expected/Value_All".Expected_81,
              Expected4 := "Expected/Value_All".Expected_82,
              Expected5 := "Expected/Value_All".Expected_83,
              Expected6 := "Expected/Value_All".Expected_84,
              Expected7 := "Expected/Value_All".Expected_85,
              Expected8 := "Expected/Value_All".Expected_86,
              Expected9 := "Expected/Value_All".Expected_87,
              Expected10 := "Expected/Value_All".Expected_88,
              Expected11 := "Expected/Value_All".Expected_89,
              Expected12 := "Expected/Value_All".Expected_90,
              Expected13 := "Expected/Value_All".Expected_91,
              Expected14 := "Expected/Value_All".Expected_92,
              Expected15 := "Expected/Value_All".Expected_93,
              Expected16 := "Expected/Value_All".Expected_94,
              Expected17 := "Expected/Value_All".Expected_95,
              Expected18 := "Expected/Value_All".Expected_96,
              Expected19 := "Expected/Value_All".Expected_97,
              Expected20 := "Expected/Value_All".Expected_98,
              Expected21 := "Expected/Value_All".Expected_99,
              Expected22 := "Expected/Value_All".Expected_100,
              Expected23 := "Expected/Value_All".Expected_101,
              Expected24 := "Expected/Value_All".Expected_102,
              Expected25 := "Expected/Value_All".Expected_103,
              Expected26 := "Expected/Value_All".Expected_104,
              On_Motor => "Output Step Motor No.4",
              ENO => #_w6);
   IF #_w6 AND "Output Step Motor No.4" THEN
       "SR_System_In Motor No.1(6)" := TRUE;   // SR flip-flop
   END_IF;
   IF "Output Motor 1,2 fower จัดเก็บ 4" THEN "SR_System_In Motor No.1(6)" := FALSE; END_IF;
   #_w9 := "SR_System_In Motor No.1(6)";
   "Expected"(Expected1 := "Expected/Value_All".Expected_105,
              Expected2 := "Expected/Value_All".Expected_106,
              Expected3 := "Expected/Value_All".Expected_107,
              Expected4 := "Expected/Value_All".Expected_108,
              Expected5 := "Expected/Value_All".Expected_109,
              Expected6 := "Expected/Value_All".Expected_110,
              Expected7 := "Expected/Value_All".Expected_111,
              Expected8 := "Expected/Value_All".Expected_112,
              Expected9 := "Expected/Value_All".Expected_113,
              Expected10 := "Expected/Value_All".Expected_114,
              Expected11 := "Expected/Value_All".Expected_115,
              Expected12 := "Expected/Value_All".Expected_116,
              Expected13 := "Expected/Value_All".Expected_117,
              Expected14 := "Expected/Value_All".Expected_118,
              Expected15 := "Expected/Value_All".Expected_119,
              Expected16 := "Expected/Value_All".Expected_120,
              Expected17 := "Expected/Value_All".Expected_121,
              Expected18 := "Expected/Value_All".Expected_122,
              Expected19 := "Expected/Value_All".Expected_123,
              Expected20 := "Expected/Value_All".Expected_124,
              Expected21 := "Expected/Value_All".Expected_125,
              Expected22 := "Expected/Value_All".Expected_126,
              Expected23 := "Expected/Value_All".Expected_127,
              Expected24 := "Expected/Value_All".Expected_128,
              Expected25 := "Expected/Value_All".Expected_129,
              Expected26 := "Expected/Value_All".Expected_130,
              On_Motor => "Output Step Motor No.5",
              ENO => #_w8);
   IF #_w8 AND "Output Step Motor No.5" THEN
       "SR_System_In Motor No.1(8)" := TRUE;   // SR flip-flop
   END_IF;
   IF "Output Motor 1,2 fower จัดเก็บ 5" THEN "SR_System_In Motor No.1(8)" := FALSE; END_IF;
   #_w11 := "SR_System_In Motor No.1(8)";
   "Expected"(Expected1 := "Expected/Value_All".Expected_131,
              Expected2 := "Expected/Value_All".Expected_132,
              Expected3 := "Expected/Value_All".Expected_133,
              Expected4 := "Expected/Value_All".Expected_134,
              Expected5 := "Expected/Value_All".Expected_135,
              Expected6 := "Expected/Value_All".Expected_136,
              Expected7 := "Expected/Value_All".Expected_137,
              Expected8 := "Expected/Value_All".Expected_138,
              Expected9 := "Expected/Value_All".Expected_139,
              Expected10 := "Expected/Value_All".Expected_140,
              Expected11 := "Expected/Value_All".Expected_141,
              Expected12 := "Expected/Value_All".Expected_142,
              Expected13 := "Expected/Value_All".Expected_143,
              Expected14 := "Expected/Value_All".Expected_144,
              Expected15 := "Expected/Value_All".Expected_145,
              Expected16 := "Expected/Value_All".Expected_146,
              Expected17 := "Expected/Value_All".Expected_147,
              Expected18 := "Expected/Value_All".Expected_148,
              Expected19 := "Expected/Value_All".Expected_149,
              Expected20 := "Expected/Value_All".Expected_150,
              Expected21 := "Expected/Value_All".Expected_151,
              Expected22 := "Expected/Value_All".Expected_152,
              Expected23 := "Expected/Value_All".Expected_153,
              Expected24 := "Expected/Value_All".Expected_154,
              Expected25 := "Expected/Value_All".Expected_155,
              Expected26 := "Expected/Value_All".Expected_156,
              On_Motor => "Output Step Motor No.6",
              ENO => #_w10);
   IF #_w10 AND "Output Step Motor No.6" THEN
       "SR_System_In Motor No.1(10)" := TRUE;   // SR flip-flop
   END_IF;
   IF "Output Motor 1,2 fower จัดเก็บ 6" THEN "SR_System_In Motor No.1(10)" := FALSE; END_IF;
   #_w13 := "SR_System_In Motor No.1(10)";
   "Expected"(Expected1 := "Expected/Value_All".Expected_157,
              Expected2 := "Expected/Value_All".Expected_158,
              Expected3 := "Expected/Value_All".Expected_159,
              Expected4 := "Expected/Value_All".Expected_160,
              Expected5 := "Expected/Value_All".Expected_161,
              Expected6 := "Expected/Value_All".Expected_162,
              Expected7 := "Expected/Value_All".Expected_163,
              Expected8 := "Expected/Value_All".Expected_164,
              Expected9 := "Expected/Value_All".Expected_165,
              Expected10 := "Expected/Value_All".Expected_166,
              Expected11 := "Expected/Value_All".Expected_167,
              Expected12 := "Expected/Value_All".Expected_168,
              Expected13 := "Expected/Value_All".Expected_169,
              Expected14 := "Expected/Value_All".Expected_170,
              Expected15 := "Expected/Value_All".Expected_171,
              Expected16 := "Expected/Value_All".Expected_172,
              Expected17 := "Expected/Value_All".Expected_173,
              Expected18 := "Expected/Value_All".Expected_174,
              Expected19 := "Expected/Value_All".Expected_175,
              Expected20 := "Expected/Value_All".Expected_176,
              Expected21 := "Expected/Value_All".Expected_177,
              Expected22 := "Expected/Value_All".Expected_178,
              Expected23 := "Expected/Value_All".Expected_179,
              Expected24 := "Expected/Value_All".Expected_180,
              Expected25 := "Expected/Value_All".Expected_181,
              Expected26 := "Expected/Value_All".Expected_182,
              On_Motor => "Output Step Motor No.7",
              ENO => #_w12);
   IF #_w12 AND "Output Step Motor No.7" THEN
       "SR_System_In Motor No.1(12)" := TRUE;   // SR flip-flop
   END_IF;
   IF "Output Motor 1,2 fower จัดเก็บ 7" THEN "SR_System_In Motor No.1(12)" := FALSE; END_IF;
   #_w15 := "SR_System_In Motor No.1(12)";
   "Expected"(Expected1 := "Expected/Value_All".Expected_183,
              Expected2 := "Expected/Value_All".Expected_184,
              Expected3 := "Expected/Value_All".Expected_185,
              Expected4 := "Expected/Value_All".Expected_186,
              Expected5 := "Expected/Value_All".Expected_187,
              Expected6 := "Expected/Value_All".Expected_188,
              Expected7 := "Expected/Value_All".Expected_189,
              Expected8 := "Expected/Value_All".Expected_190,
              Expected9 := "Expected/Value_All".Expected_191,
              Expected10 := "Expected/Value_All".Expected_192,
              Expected11 := "Expected/Value_All".Expected_193,
              Expected12 := "Expected/Value_All".Expected_194,
              Expected13 := "Expected/Value_All".Expected_195,
              Expected14 := "Expected/Value_All".Expected_196,
              Expected15 := "Expected/Value_All".Expected_197,
              Expected16 := "Expected/Value_All".Expected_198,
              Expected17 := "Expected/Value_All".Expected_199,
              Expected18 := "Expected/Value_All".Expected_200,
              Expected19 := "Expected/Value_All".Expected_201,
              Expected20 := "Expected/Value_All".Expected_202,
              Expected21 := "Expected/Value_All".Expected_203,
              Expected22 := "Expected/Value_All".Expected_204,
              Expected23 := "Expected/Value_All".Expected_205,
              Expected24 := "Expected/Value_All".Expected_206,
              Expected25 := "Expected/Value_All".Expected_207,
              Expected26 := "Expected/Value_All".Expected_208,
              On_Motor => "Output Step Motor No.8",
              ENO => #_w14);
   IF #_w14 AND "Output Step Motor No.8" THEN
       "SR_System_In Motor No.1(14)" := TRUE;   // SR flip-flop
   END_IF;
   IF "Output Motor 1,2 fower จัดเก็บ 8" THEN "SR_System_In Motor No.1(14)" := FALSE; END_IF;
   #_w17 := "SR_System_In Motor No.1(14)";
   "Expected"(Expected1 := "Expected/Value_All".Expected_209,
              Expected2 := "Expected/Value_All".Expected_210,
              Expected3 := "Expected/Value_All".Expected_211,
              Expected4 := "Expected/Value_All".Expected_212,
              Expected5 := "Expected/Value_All".Expected_213,
              Expected6 := "Expected/Value_All".Expected_214,
              Expected7 := "Expected/Value_All".Expected_215,
              Expected8 := "Expected/Value_All".Expected_216,
              Expected9 := "Expected/Value_All".Expected_217,
              Expected10 := "Expected/Value_All".Expected_218,
              Expected11 := "Expected/Value_All".Expected_219,
              Expected12 := "Expected/Value_All".Expected_220,
              Expected13 := "Expected/Value_All".Expected_221,
              Expected14 := "Expected/Value_All".Expected_222,
              Expected15 := "Expected/Value_All".Expected_223,
              Expected16 := "Expected/Value_All".Expected_224,
              Expected17 := "Expected/Value_All".Expected_225,
              Expected18 := "Expected/Value_All".Expected_226,
              Expected19 := "Expected/Value_All".Expected_227,
              Expected20 := "Expected/Value_All".Expected_228,
              Expected21 := "Expected/Value_All".Expected_229,
              Expected22 := "Expected/Value_All".Expected_230,
              Expected23 := "Expected/Value_All".Expected_231,
              Expected24 := "Expected/Value_All".Expected_232,
              Expected25 := "Expected/Value_All".Expected_233,
              Expected26 := "Expected/Value_All".Expected_234,
              On_Motor => "Output Step Motor No.9",
              ENO => #_w16);
   IF #_w16 AND "Output Step Motor No.9" THEN
       "SR_System_In Motor No.1(16)" := TRUE;   // SR flip-flop
   END_IF;
   IF "Output Motor 1,2 fower จัดเก็บ 9" THEN "SR_System_In Motor No.1(16)" := FALSE; END_IF;
   #_w19 := "SR_System_In Motor No.1(16)";
   "Expected"(Expected1 := "Expected/Value_All".Expected_235,
              Expected2 := "Expected/Value_All".Expected_236,
              Expected3 := "Expected/Value_All".Expected_237,
              Expected4 := "Expected/Value_All".Expected_238,
              Expected5 := "Expected/Value_All".Expected_239,
              Expected6 := "Expected/Value_All".Expected_240,
              Expected7 := "Expected/Value_All".Expected_241,
              Expected8 := "Expected/Value_All".Expected_242,
              Expected9 := "Expected/Value_All".Expected_243,
              Expected10 := "Expected/Value_All".Expected_244,
              Expected11 := "Expected/Value_All".Expected_245,
              Expected12 := "Expected/Value_All".Expected_246,
              Expected13 := "Expected/Value_All".Expected_247,
              Expected14 := "Expected/Value_All".Expected_248,
              Expected15 := "Expected/Value_All".Expected_249,
              Expected16 := "Expected/Value_All".Expected_250,
              Expected17 := "Expected/Value_All".Expected_251,
              Expected18 := "Expected/Value_All".Expected_252,
              Expected19 := "Expected/Value_All".Expected_253,
              Expected20 := "Expected/Value_All".Expected_254,
              Expected21 := "Expected/Value_All".Expected_255,
              Expected22 := "Expected/Value_All".Expected_256,
              Expected23 := "Expected/Value_All".Expected_257,
              Expected24 := "Expected/Value_All".Expected_258,
              Expected25 := "Expected/Value_All".Expected_259,
              Expected26 := "Expected/Value_All".Expected_260,
              On_Motor => "Output Step Motor No.10",
              ENO => #_w18);
   IF #_w18 AND "Output Step Motor No.10" THEN
       "SR_System_In Motor No.1(18)" := TRUE;   // SR flip-flop
   END_IF;
   IF "Output Motor 1,2 fower จัดเก็บ 10" THEN "SR_System_In Motor No.1(18)" := FALSE; END_IF;
   #_w21 := "SR_System_In Motor No.1(18)";
   "Expected"(Expected1 := "Expected/Value_All".Expected_261,
              Expected2 := "Expected/Value_All".Expected_262,
              Expected3 := "Expected/Value_All".Expected_263,
              Expected4 := "Expected/Value_All".Expected_264,
              Expected5 := "Expected/Value_All".Expected_265,
              Expected6 := "Expected/Value_All".Expected_266,
              Expected7 := "Expected/Value_All".Expected_267,
              Expected8 := "Expected/Value_All".Expected_268,
              Expected9 := "Expected/Value_All".Expected_269,
              Expected10 := "Expected/Value_All".Expected_270,
              Expected11 := "Expected/Value_All".Expected_271,
              Expected12 := "Expected/Value_All".Expected_272,
              Expected13 := "Expected/Value_All".Expected_273,
              Expected14 := "Expected/Value_All".Expected_274,
              Expected15 := "Expected/Value_All".Expected_275,
              Expected16 := "Expected/Value_All".Expected_276,
              Expected17 := "Expected/Value_All".Expected_277,
              Expected18 := "Expected/Value_All".Expected_278,
              Expected19 := "Expected/Value_All".Expected_279,
              Expected20 := "Expected/Value_All".Expected_280,
              Expected21 := "Expected/Value_All".Expected_281,
              Expected22 := "Expected/Value_All".Expected_282,
              Expected23 := "Expected/Value_All".Expected_283,
              Expected24 := "Expected/Value_All".Expected_284,
              Expected25 := "Expected/Value_All".Expected_285,
              Expected26 := "Expected/Value_All".Expected_286,
              On_Motor => "Output Step Motor No.11",
              ENO => #_w20);
   IF #_w20 AND "Output Step Motor No.11" THEN
       "SR_System_In Motor No.1(20)" := TRUE;   // SR flip-flop
   END_IF;
   IF "Output Motor 1,2 fower จัดเก็บ 11" THEN "SR_System_In Motor No.1(20)" := FALSE; END_IF;
   #_w23 := "SR_System_In Motor No.1(20)";
   "Expected"(Expected1 := "Expected/Value_All".Expected_287,
              Expected2 := "Expected/Value_All".Expected_288,
              Expected3 := "Expected/Value_All".Expected_289,
              Expected4 := "Expected/Value_All".Expected_290,
              Expected5 := "Expected/Value_All".Expected_291,
              Expected6 := "Expected/Value_All".Expected_292,
              Expected7 := "Expected/Value_All".Expected_293,
              Expected8 := "Expected/Value_All".Expected_294,
              Expected9 := "Expected/Value_All".Expected_295,
              Expected10 := "Expected/Value_All".Expected_296,
              Expected11 := "Expected/Value_All".Expected_297,
              Expected12 := "Expected/Value_All".Expected_298,
              Expected13 := "Expected/Value_All".Expected_299,
              Expected14 := "Expected/Value_All".Expected_300,
              Expected15 := "Expected/Value_All".Expected_301,
              Expected16 := "Expected/Value_All".Expected_302,
              Expected17 := "Expected/Value_All".Expected_303,
              Expected18 := "Expected/Value_All".Expected_304,
              Expected19 := "Expected/Value_All".Expected_305,
              Expected20 := "Expected/Value_All".Expected_306,
              Expected21 := "Expected/Value_All".Expected_307,
              Expected22 := "Expected/Value_All".Expected_308,
              Expected23 := "Expected/Value_All".Expected_309,
              Expected24 := "Expected/Value_All".Expected_310,
              Expected25 := "Expected/Value_All".Expected_311,
              Expected26 := "Expected/Value_All".Expected_312,
              On_Motor => "Output Step Motor No.12",
              ENO => #_w22);
   IF #_w22 AND "Output Step Motor No.12" THEN
       "SR_System_In Motor No.1(22)" := TRUE;   // SR flip-flop
   END_IF;
   IF "Output Motor 1,2 fower จัดเก็บ 12" THEN "SR_System_In Motor No.1(22)" := FALSE; END_IF;
   #_w25 := "SR_System_In Motor No.1(22)";
   "Expected"(Expected1 := "Expected/Value_All".Expected_313,
              Expected2 := "Expected/Value_All".Expected_314,
              Expected3 := "Expected/Value_All".Expected_315,
              Expected4 := "Expected/Value_All".Expected_316,
              Expected5 := "Expected/Value_All".Expected_317,
              Expected6 := "Expected/Value_All".Expected_318,
              Expected7 := "Expected/Value_All".Expected_319,
              Expected8 := "Expected/Value_All".Expected_320,
              Expected9 := "Expected/Value_All".Expected_321,
              Expected10 := "Expected/Value_All".Expected_322,
              Expected11 := "Expected/Value_All".Expected_323,
              Expected12 := "Expected/Value_All".Expected_324,
              Expected13 := "Expected/Value_All".Expected_325,
              Expected14 := "Expected/Value_All".Expected_326,
              Expected15 := "Expected/Value_All".Expected_327,
              Expected16 := "Expected/Value_All".Expected_328,
              Expected17 := "Expected/Value_All".Expected_329,
              Expected18 := "Expected/Value_All".Expected_330,
              Expected19 := "Expected/Value_All".Expected_331,
              Expected20 := "Expected/Value_All".Expected_332,
              Expected21 := "Expected/Value_All".Expected_333,
              Expected22 := "Expected/Value_All".Expected_334,
              Expected23 := "Expected/Value_All".Expected_335,
              Expected24 := "Expected/Value_All".Expected_336,
              Expected25 := "Expected/Value_All".Expected_337,
              Expected26 := "Expected/Value_All".Expected_338,
              On_Motor => "Output Step Motor No.13",
              ENO => #_w24);
   IF #_w24 AND "Output Step Motor No.13" THEN
       "SR_System_In Motor No.1(24)" := TRUE;   // SR flip-flop
   END_IF;
   IF "Output Motor 1,2 fower จัดเก็บ 13" THEN "SR_System_In Motor No.1(24)" := FALSE; END_IF;
   #_w27 := "SR_System_In Motor No.1(24)";
   "Expected"(Expected1 := "Expected/Value_All".Expected_339,
              Expected2 := "Expected/Value_All".Expected_340,
              Expected3 := "Expected/Value_All".Expected_341,
              Expected4 := "Expected/Value_All".Expected_342,
              Expected5 := "Expected/Value_All".Expected_343,
              Expected6 := "Expected/Value_All".Expected_344,
              Expected7 := "Expected/Value_All".Expected_345,
              Expected8 := "Expected/Value_All".Expected_346,
              Expected9 := "Expected/Value_All".Expected_347,
              Expected10 := "Expected/Value_All".Expected_348,
              Expected11 := "Expected/Value_All".Expected_349,
              Expected12 := "Expected/Value_All".Expected_350,
              Expected13 := "Expected/Value_All".Expected_351,
              Expected14 := "Expected/Value_All".Expected_352,
              Expected15 := "Expected/Value_All".Expected_353,
              Expected16 := "Expected/Value_All".Expected_354,
              Expected17 := "Expected/Value_All".Expected_355,
              Expected18 := "Expected/Value_All".Expected_356,
              Expected19 := "Expected/Value_All".Expected_357,
              Expected20 := "Expected/Value_All".Expected_358,
              Expected21 := "Expected/Value_All".Expected_359,
              Expected22 := "Expected/Value_All".Expected_360,
              Expected23 := "Expected/Value_All".Expected_361,
              Expected24 := "Expected/Value_All".Expected_362,
              Expected25 := "Expected/Value_All".Expected_363,
              Expected26 := "Expected/Value_All".Expected_364,
              On_Motor => "Output Step Motor No.14",
              ENO => #_w26);
   IF #_w26 AND "Output Step Motor No.14" THEN
       "SR_System_In Motor No.1(26)" := TRUE;   // SR flip-flop
   END_IF;
   IF "Output Motor 1,2 fower จัดเก็บ 14" THEN "SR_System_In Motor No.1(26)" := FALSE; END_IF;
   #_w29 := "SR_System_In Motor No.1(26)";
   "Expected"(Expected1 := "Expected/Value_All".Expected_365,
              Expected2 := "Expected/Value_All".Expected_366,
              Expected3 := "Expected/Value_All".Expected_367,
              Expected4 := "Expected/Value_All".Expected_368,
              Expected5 := "Expected/Value_All".Expected_369,
              Expected6 := "Expected/Value_All".Expected_370,
              Expected7 := "Expected/Value_All".Expected_371,
              Expected8 := "Expected/Value_All".Expected_372,
              Expected9 := "Expected/Value_All".Expected_373,
              Expected10 := "Expected/Value_All".Expected_374,
              Expected11 := "Expected/Value_All".Expected_375,
              Expected12 := "Expected/Value_All".Expected_376,
              Expected13 := "Expected/Value_All".Expected_377,
              Expected14 := "Expected/Value_All".Expected_378,
              Expected15 := "Expected/Value_All".Expected_379,
              Expected16 := "Expected/Value_All".Expected_380,
              Expected17 := "Expected/Value_All".Expected_381,
              Expected18 := "Expected/Value_All".Expected_382,
              Expected19 := "Expected/Value_All".Expected_383,
              Expected20 := "Expected/Value_All".Expected_384,
              Expected21 := "Expected/Value_All".Expected_385,
              Expected22 := "Expected/Value_All".Expected_386,
              Expected23 := "Expected/Value_All".Expected_387,
              Expected24 := "Expected/Value_All".Expected_388,
              Expected25 := "Expected/Value_All".Expected_389,
              Expected26 := "Expected/Value_All".Expected_390,
              On_Motor => "Output Step Motor No.15",
              ENO => #_w28);
   IF #_w28 AND "Output Step Motor No.15" THEN
       "SR_System_In Motor No.1(28)" := TRUE;   // SR flip-flop
   END_IF;
   IF "Output Motor 1,2 fower จัดเก็บ 15" THEN "SR_System_In Motor No.1(28)" := FALSE; END_IF;
   #_w31 := "SR_System_In Motor No.1(28)";
   "Expected"(Expected1 := "Expected/Value_All".Expected_391,
              Expected2 := "Expected/Value_All".Expected_392,
              Expected3 := "Expected/Value_All".Expected_393,
              Expected4 := "Expected/Value_All".Expected_394,
              Expected5 := "Expected/Value_All".Expected_395,
              Expected6 := "Expected/Value_All".Expected_396,
              Expected7 := "Expected/Value_All".Expected_397,
              Expected8 := "Expected/Value_All".Expected_398,
              Expected9 := "Expected/Value_All".Expected_399,
              Expected10 := "Expected/Value_All".Expected_400,
              Expected11 := "Expected/Value_All".Expected_401,
              Expected12 := "Expected/Value_All".Expected_402,
              Expected13 := "Expected/Value_All".Expected_403,
              Expected14 := "Expected/Value_All".Expected_404,
              Expected15 := "Expected/Value_All".Expected_405,
              Expected16 := "Expected/Value_All".Expected_406,
              Expected17 := "Expected/Value_All".Expected_407,
              Expected18 := "Expected/Value_All".Expected_408,
              Expected19 := "Expected/Value_All".Expected_409,
              Expected20 := "Expected/Value_All".Expected_410,
              Expected21 := "Expected/Value_All".Expected_411,
              Expected22 := "Expected/Value_All".Expected_412,
              Expected23 := "Expected/Value_All".Expected_413,
              Expected24 := "Expected/Value_All".Expected_414,
              Expected25 := "Expected/Value_All".Expected_415,
              Expected26 := "Expected/Value_All".Expected_416,
              On_Motor => "Output Step Motor No.16",
              ENO => #_w30);
   IF #_w30 AND "Output Step Motor No.16" THEN
       "SR_System_In Motor No.1(30)" := TRUE;   // SR flip-flop
   END_IF;
   IF "Output Motor 1,2 fower จัดเก็บ 16" THEN "SR_System_In Motor No.1(30)" := FALSE; END_IF;
   #_w33 := "SR_System_In Motor No.1(30)";
   "Expected"(Expected1 := "Expected/Value_All".Expected_417,
              Expected2 := "Expected/Value_All".Expected_418,
              Expected3 := "Expected/Value_All".Expected_419,
              Expected4 := "Expected/Value_All".Expected_420,
              Expected5 := "Expected/Value_All".Expected_421,
              Expected6 := "Expected/Value_All".Expected_422,
              Expected7 := "Expected/Value_All".Expected_423,
              Expected8 := "Expected/Value_All".Expected_424,
              Expected9 := "Expected/Value_All".Expected_425,
              Expected10 := "Expected/Value_All".Expected_426,
              Expected11 := "Expected/Value_All".Expected_427,
              Expected12 := "Expected/Value_All".Expected_428,
              Expected13 := "Expected/Value_All".Expected_429,
              Expected14 := "Expected/Value_All".Expected_430,
              Expected15 := "Expected/Value_All".Expected_431,
              Expected16 := "Expected/Value_All".Expected_432,
              Expected17 := "Expected/Value_All".Expected_433,
              Expected18 := "Expected/Value_All".Expected_434,
              Expected19 := "Expected/Value_All".Expected_435,
              Expected20 := "Expected/Value_All".Expected_436,
              Expected21 := "Expected/Value_All".Expected_437,
              Expected22 := "Expected/Value_All".Expected_438,
              Expected23 := "Expected/Value_All".Expected_439,
              Expected24 := "Expected/Value_All".Expected_440,
              Expected25 := "Expected/Value_All".Expected_441,
              Expected26 := "Expected/Value_All".Expected_442,
              On_Motor => "Output Step Motor No.17",
              ENO => #_w32);
   IF #_w32 AND "Output Step Motor No.17" THEN
       "SR_System_In Motor No.1(32)" := TRUE;   // SR flip-flop
   END_IF;
   IF "Output Motor 1,2 fower จัดเก็บ 17" THEN "SR_System_In Motor No.1(32)" := FALSE; END_IF;
   #_w35 := "SR_System_In Motor No.1(32)";
   "Expected"(Expected1 := "Expected/Value_All".Expected_443,
              Expected2 := "Expected/Value_All".Expected_444,
              Expected3 := "Expected/Value_All".Expected_445,
              Expected4 := "Expected/Value_All".Expected_446,
              Expected5 := "Expected/Value_All".Expected_447,
              Expected6 := "Expected/Value_All".Expected_448,
              Expected7 := "Expected/Value_All".Expected_449,
              Expected8 := "Expected/Value_All".Expected_450,
              Expected9 := "Expected/Value_All".Expected_451,
              Expected10 := "Expected/Value_All".Expected_452,
              Expected11 := "Expected/Value_All".Expected_453,
              Expected12 := "Expected/Value_All".Expected_454,
              Expected13 := "Expected/Value_All".Expected_455,
              Expected14 := "Expected/Value_All".Expected_456,
              Expected15 := "Expected/Value_All".Expected_457,
              Expected16 := "Expected/Value_All".Expected_458,
              Expected17 := "Expected/Value_All".Expected_459,
              Expected18 := "Expected/Value_All".Expected_460,
              Expected19 := "Expected/Value_All".Expected_461,
              Expected20 := "Expected/Value_All".Expected_462,
              Expected21 := "Expected/Value_All".Expected_463,
              Expected22 := "Expected/Value_All".Expected_464,
              Expected23 := "Expected/Value_All".Expected_465,
              Expected24 := "Expected/Value_All".Expected_466,
              Expected25 := "Expected/Value_All".Expected_467,
              Expected26 := "Expected/Value_All".Expected_468,
              On_Motor => "Output Step Motor No.18",
              ENO => #_w34);
   IF #_w34 AND "Output Step Motor No.18" THEN
       "SR_System_In Motor No.1(34)" := TRUE;   // SR flip-flop
   END_IF;
   IF "Output Motor 1,2 fower จัดเก็บ 18" THEN "SR_System_In Motor No.1(34)" := FALSE; END_IF;
   #_w37 := "SR_System_In Motor No.1(34)";
   "Expected"(Expected1 := "Expected/Value_All".Expected_469,
              Expected2 := "Expected/Value_All".Expected_470,
              Expected3 := "Expected/Value_All".Expected_471,
              Expected4 := "Expected/Value_All".Expected_472,
              Expected5 := "Expected/Value_All".Expected_473,
              Expected6 := "Expected/Value_All".Expected_474,
              Expected7 := "Expected/Value_All".Expected_475,
              Expected8 := "Expected/Value_All".Expected_476,
              Expected9 := "Expected/Value_All".Expected_477,
              Expected10 := "Expected/Value_All".Expected_478,
              Expected11 := "Expected/Value_All".Expected_479,
              Expected12 := "Expected/Value_All".Expected_480,
              Expected13 := "Expected/Value_All".Expected_481,
              Expected14 := "Expected/Value_All".Expected_482,
              Expected15 := "Expected/Value_All".Expected_483,
              Expected16 := "Expected/Value_All".Expected_484,
              Expected17 := "Expected/Value_All".Expected_485,
              Expected18 := "Expected/Value_All".Expected_486,
              Expected19 := "Expected/Value_All".Expected_487,
              Expected20 := "Expected/Value_All".Expected_488,
              Expected21 := "Expected/Value_All".Expected_489,
              Expected22 := "Expected/Value_All".Expected_490,
              Expected23 := "Expected/Value_All".Expected_491,
              Expected24 := "Expected/Value_All".Expected_492,
              Expected25 := "Expected/Value_All".Expected_493,
              Expected26 := "Expected/Value_All".Expected_494,
              On_Motor => "Output Step Motor No.19",
              ENO => #_w36);
   IF #_w36 AND "Output Step Motor No.19" THEN
       "SR_System_In Motor No.1(36)" := TRUE;   // SR flip-flop
   END_IF;
   IF "Output Motor 1,2 fower จัดเก็บ 19" THEN "SR_System_In Motor No.1(36)" := FALSE; END_IF;
   #_w39 := "SR_System_In Motor No.1(36)";
   "Expected"(Expected1 := "Expected/Value_All".Expected_495,
              Expected2 := "Expected/Value_All".Expected_496,
              Expected3 := "Expected/Value_All".Expected_497,
              Expected4 := "Expected/Value_All".Expected_498,
              Expected5 := "Expected/Value_All".Expected_499,
              Expected6 := "Expected/Value_All".Expected_500,
              Expected7 := "Expected/Value_All".Expected_501,
              Expected8 := "Expected/Value_All".Expected_502,
              Expected9 := "Expected/Value_All".Expected_503,
              Expected10 := "Expected/Value_All".Expected_504,
              Expected11 := "Expected/Value_All".Expected_505,
              Expected12 := "Expected/Value_All".Expected_506,
              Expected13 := "Expected/Value_All".Expected_507,
              Expected14 := "Expected/Value_All".Expected_508,
              Expected15 := "Expected/Value_All".Expected_509,
              Expected16 := "Expected/Value_All".Expected_510,
              Expected17 := "Expected/Value_All".Expected_511,
              Expected18 := "Expected/Value_All".Expected_512,
              Expected19 := "Expected/Value_All".Expected_513,
              Expected20 := "Expected/Value_All".Expected_514,
              Expected21 := "Expected/Value_All".Expected_515,
              Expected22 := "Expected/Value_All".Expected_516,
              Expected23 := "Expected/Value_All".Expected_517,
              Expected24 := "Expected/Value_All".Expected_518,
              Expected25 := "Expected/Value_All".Expected_519,
              Expected26 := "Expected/Value_All".Expected_520,
              On_Motor => "Output Step Motor No.20",
              ENO => #_w38);
   IF #_w38 AND "Output Step Motor No.20" THEN
       "SR_System_In Motor No.1(38)" := TRUE;   // SR flip-flop
   END_IF;
   IF "Output Motor 1,2 fower จัดเก็บ 20" THEN "SR_System_In Motor No.1(38)" := FALSE; END_IF;
   "test หลังเคลื่อนที่มาตำแหน่งปล่อยกล่องยา"(EN := #_w3 OR #_w5 OR #_w7 OR #_w9 OR #_w11 OR #_w13 OR #_w15 OR #_w17 OR #_w19 OR #_w21 OR #_w23 OR #_w25 OR #_w27 OR #_w29 OR #_w31 OR #_w33 OR #_w35 OR #_w37 OR #_w39 OR "SR_System_In Motor No.1(38)",
                           ENO => #_w40);
   #"Stepper Motor  ทำงาน" := #_w40 AND "หมุนไปตำแหต่งปล่อยกล่องยา";
END_REGION

REGION Network 2
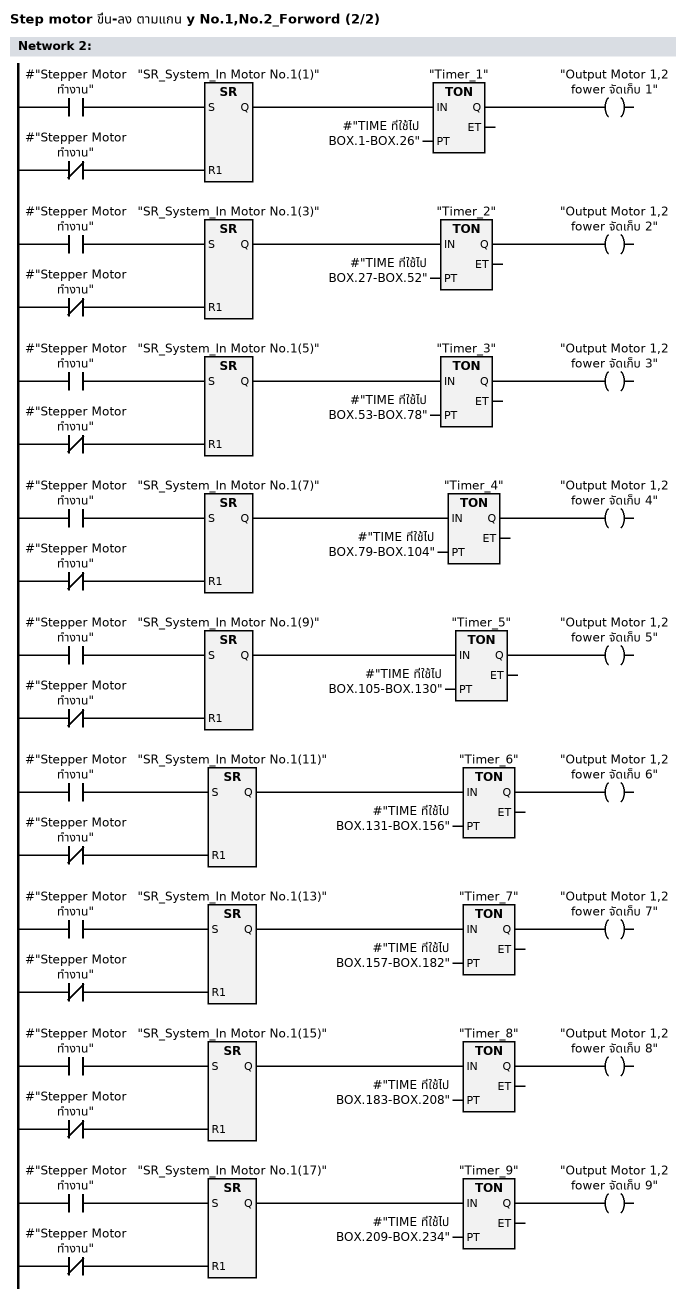
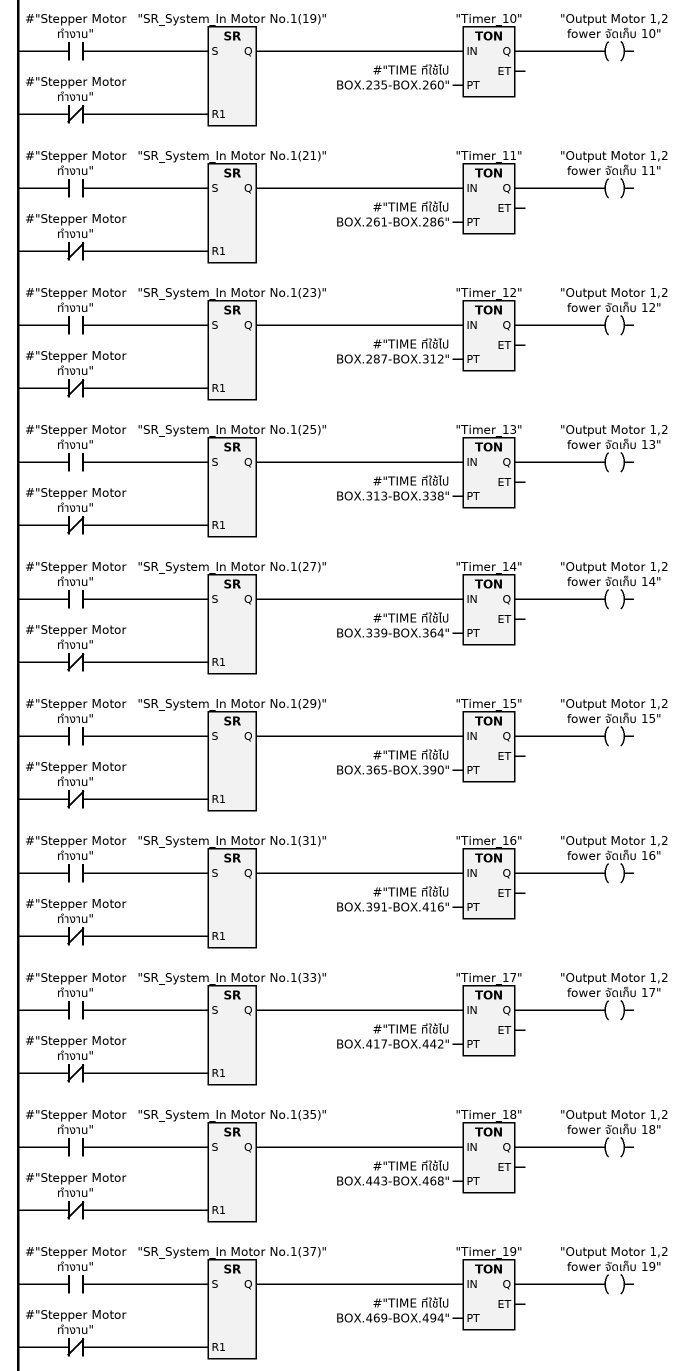
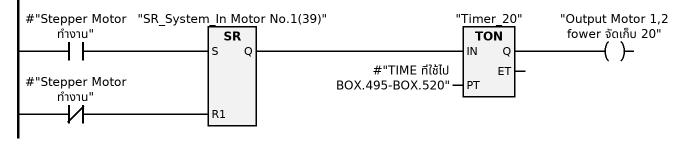
   IF #"Stepper Motor  ทำงาน" THEN
       "SR_System_In Motor No.1(1)" := TRUE;   // SR flip-flop
   END_IF;
   IF NOT #"Stepper Motor  ทำงาน" THEN "SR_System_In Motor No.1(1)" := FALSE; END_IF;
   "Timer_1".TON(IN := "SR_System_In Motor No.1(1)", PT := #"TIME ที่ใช้ไป BOX.1-BOX.26");
   "Output Motor 1,2 fower จัดเก็บ 1" := "Timer_1".Q;
   IF #"Stepper Motor  ทำงาน" THEN
       "SR_System_In Motor No.1(3)" := TRUE;   // SR flip-flop
   END_IF;
   IF NOT #"Stepper Motor  ทำงาน" THEN "SR_System_In Motor No.1(3)" := FALSE; END_IF;
   "Timer_2".TON(IN := "SR_System_In Motor No.1(3)", PT := #"TIME ที่ใช้ไป BOX.27-BOX.52");
   "Output Motor 1,2 fower จัดเก็บ 2" := "Timer_2".Q;
   IF #"Stepper Motor  ทำงาน" THEN
       "SR_System_In Motor No.1(5)" := TRUE;   // SR flip-flop
   END_IF;
   IF NOT #"Stepper Motor  ทำงาน" THEN "SR_System_In Motor No.1(5)" := FALSE; END_IF;
   "Timer_3".TON(IN := "SR_System_In Motor No.1(5)", PT := #"TIME ที่ใช้ไป BOX.53-BOX.78");
   "Output Motor 1,2 fower จัดเก็บ 3" := "Timer_3".Q;
   IF #"Stepper Motor  ทำงาน" THEN
       "SR_System_In Motor No.1(7)" := TRUE;   // SR flip-flop
   END_IF;
   IF NOT #"Stepper Motor  ทำงาน" THEN "SR_System_In Motor No.1(7)" := FALSE; END_IF;
   "Timer_4".TON(IN := "SR_System_In Motor No.1(7)", PT := #"TIME ที่ใช้ไป BOX.79-BOX.104");
   "Output Motor 1,2 fower จัดเก็บ 4" := "Timer_4".Q;
   IF #"Stepper Motor  ทำงาน" THEN
       "SR_System_In Motor No.1(9)" := TRUE;   // SR flip-flop
   END_IF;
   IF NOT #"Stepper Motor  ทำงาน" THEN "SR_System_In Motor No.1(9)" := FALSE; END_IF;
   "Timer_5".TON(IN := "SR_System_In Motor No.1(9)", PT := #"TIME ที่ใช้ไป BOX.105-BOX.130");
   "Output Motor 1,2 fower จัดเก็บ 5" := "Timer_5".Q;
   IF #"Stepper Motor  ทำงาน" THEN
       "SR_System_In Motor No.1(11)" := TRUE;   // SR flip-flop
   END_IF;
   IF NOT #"Stepper Motor  ทำงาน" THEN "SR_System_In Motor No.1(11)" := FALSE; END_IF;
   "Timer_6".TON(IN := "SR_System_In Motor No.1(11)", PT := #"TIME ที่ใช้ไป BOX.131-BOX.156");
   "Output Motor 1,2 fower จัดเก็บ 6" := "Timer_6".Q;
   IF #"Stepper Motor  ทำงาน" THEN
       "SR_System_In Motor No.1(13)" := TRUE;   // SR flip-flop
   END_IF;
   IF NOT #"Stepper Motor  ทำงาน" THEN "SR_System_In Motor No.1(13)" := FALSE; END_IF;
   "Timer_7".TON(IN := "SR_System_In Motor No.1(13)", PT := #"TIME ที่ใช้ไป BOX.157-BOX.182");
   "Output Motor 1,2 fower จัดเก็บ 7" := "Timer_7".Q;
   IF #"Stepper Motor  ทำงาน" THEN
       "SR_System_In Motor No.1(15)" := TRUE;   // SR flip-flop
   END_IF;
   IF NOT #"Stepper Motor  ทำงาน" THEN "SR_System_In Motor No.1(15)" := FALSE; END_IF;
   "Timer_8".TON(IN := "SR_System_In Motor No.1(15)", PT := #"TIME ที่ใช้ไป BOX.183-BOX.208");
   "Output Motor 1,2 fower จัดเก็บ 8" := "Timer_8".Q;
   IF #"Stepper Motor  ทำงาน" THEN
       "SR_System_In Motor No.1(17)" := TRUE;   // SR flip-flop
   END_IF;
   IF NOT #"Stepper Motor  ทำงาน" THEN "SR_System_In Motor No.1(17)" := FALSE; END_IF;
   "Timer_9".TON(IN := "SR_System_In Motor No.1(17)", PT := #"TIME ที่ใช้ไป BOX.209-BOX.234");
   "Output Motor 1,2 fower จัดเก็บ 9" := "Timer_9".Q;
   IF #"Stepper Motor  ทำงาน" THEN
       "SR_System_In Motor No.1(19)" := TRUE;   // SR flip-flop
   END_IF;
   IF NOT #"Stepper Motor  ทำงาน" THEN "SR_System_In Motor No.1(19)" := FALSE; END_IF;
   "Timer_10".TON(IN := "SR_System_In Motor No.1(19)", PT := #"TIME ที่ใช้ไป BOX.235-BOX.260");
   "Output Motor 1,2 fower จัดเก็บ 10" := "Timer_10".Q;
   IF #"Stepper Motor  ทำงาน" THEN
       "SR_System_In Motor No.1(21)" := TRUE;   // SR flip-flop
   END_IF;
   IF NOT #"Stepper Motor  ทำงาน" THEN "SR_System_In Motor No.1(21)" := FALSE; END_IF;
   "Timer_11".TON(IN := "SR_System_In Motor No.1(21)", PT := #"TIME ที่ใช้ไป BOX.261-BOX.286");
   "Output Motor 1,2 fower จัดเก็บ 11" := "Timer_11".Q;
   IF #"Stepper Motor  ทำงาน" THEN
       "SR_System_In Motor No.1(23)" := TRUE;   // SR flip-flop
   END_IF;
   IF NOT #"Stepper Motor  ทำงาน" THEN "SR_System_In Motor No.1(23)" := FALSE; END_IF;
   "Timer_12".TON(IN := "SR_System_In Motor No.1(23)", PT := #"TIME ที่ใช้ไป BOX.287-BOX.312");
   "Output Motor 1,2 fower จัดเก็บ 12" := "Timer_12".Q;
   IF #"Stepper Motor  ทำงาน" THEN
       "SR_System_In Motor No.1(25)" := TRUE;   // SR flip-flop
   END_IF;
   IF NOT #"Stepper Motor  ทำงาน" THEN "SR_System_In Motor No.1(25)" := FALSE; END_IF;
   "Timer_13".TON(IN := "SR_System_In Motor No.1(25)", PT := #"TIME ที่ใช้ไป BOX.313-BOX.338");
   "Output Motor 1,2 fower จัดเก็บ 13" := "Timer_13".Q;
   IF #"Stepper Motor  ทำงาน" THEN
       "SR_System_In Motor No.1(27)" := TRUE;   // SR flip-flop
   END_IF;
   IF NOT #"Stepper Motor  ทำงาน" THEN "SR_System_In Motor No.1(27)" := FALSE; END_IF;
   "Timer_14".TON(IN := "SR_System_In Motor No.1(27)", PT := #"TIME ที่ใช้ไป BOX.339-BOX.364");
   "Output Motor 1,2 fower จัดเก็บ 14" := "Timer_14".Q;
   IF #"Stepper Motor  ทำงาน" THEN
       "SR_System_In Motor No.1(29)" := TRUE;   // SR flip-flop
   END_IF;
   IF NOT #"Stepper Motor  ทำงาน" THEN "SR_System_In Motor No.1(29)" := FALSE; END_IF;
   "Timer_15".TON(IN := "SR_System_In Motor No.1(29)", PT := #"TIME ที่ใช้ไป BOX.365-BOX.390");
   "Output Motor 1,2 fower จัดเก็บ 15" := "Timer_15".Q;
   IF #"Stepper Motor  ทำงาน" THEN
       "SR_System_In Motor No.1(31)" := TRUE;   // SR flip-flop
   END_IF;
   IF NOT #"Stepper Motor  ทำงาน" THEN "SR_System_In Motor No.1(31)" := FALSE; END_IF;
   "Timer_16".TON(IN := "SR_System_In Motor No.1(31)", PT := #"TIME ที่ใช้ไป BOX.391-BOX.416");
   "Output Motor 1,2 fower จัดเก็บ 16" := "Timer_16".Q;
   IF #"Stepper Motor  ทำงาน" THEN
       "SR_System_In Motor No.1(33)" := TRUE;   // SR flip-flop
   END_IF;
   IF NOT #"Stepper Motor  ทำงาน" THEN "SR_System_In Motor No.1(33)" := FALSE; END_IF;
   "Timer_17".TON(IN := "SR_System_In Motor No.1(33)", PT := #"TIME ที่ใช้ไป BOX.417-BOX.442");
   "Output Motor 1,2 fower จัดเก็บ 17" := "Timer_17".Q;
   IF #"Stepper Motor  ทำงาน" THEN
       "SR_System_In Motor No.1(35)" := TRUE;   // SR flip-flop
   END_IF;
   IF NOT #"Stepper Motor  ทำงาน" THEN "SR_System_In Motor No.1(35)" := FALSE; END_IF;
   "Timer_18".TON(IN := "SR_System_In Motor No.1(35)", PT := #"TIME ที่ใช้ไป BOX.443-BOX.468");
   "Output Motor 1,2 fower จัดเก็บ 18" := "Timer_18".Q;
   IF #"Stepper Motor  ทำงาน" THEN
       "SR_System_In Motor No.1(37)" := TRUE;   // SR flip-flop
   END_IF;
   IF NOT #"Stepper Motor  ทำงาน" THEN "SR_System_In Motor No.1(37)" := FALSE; END_IF;
   "Timer_19".TON(IN := "SR_System_In Motor No.1(37)", PT := #"TIME ที่ใช้ไป BOX.469-BOX.494");
   "Output Motor 1,2 fower จัดเก็บ 19" := "Timer_19".Q;
   IF #"Stepper Motor  ทำงาน" THEN
       "SR_System_In Motor No.1(39)" := TRUE;   // SR flip-flop
   END_IF;
   IF NOT #"Stepper Motor  ทำงาน" THEN "SR_System_In Motor No.1(39)" := FALSE; END_IF;
   "Timer_20".TON(IN := "SR_System_In Motor No.1(39)", PT := #"TIME ที่ใช้ไป BOX.495-BOX.520");
   "Output Motor 1,2 fower จัดเก็บ 20" := "Timer_20".Q;
END_REGION
END_FUNCTION_BLOCK

FUNCTION_BLOCK "Step motor ขึ่น-ลง ตามแกน y No.1_Blackword"   // FB4, LAD
{ S7_Optimized_Access := 'TRUE' }
VERSION : 0.1
   VAR_INPUT
      "เวลาเคลื่อนที่ของ Stepper Motor1จาก Box1_Backword" : Time;
      "เวลาเคลื่อนที่ของ Stepper Motor1จาก Box2_Backword" : Time;
      "เวลาเคลื่อนที่ของ Stepper Motor1จาก Box3_Backword" : Time;
      "เวลาเคลื่อนที่ของ Stepper Motor1จาก Box4_Backword" : Time;
      "เวลาเคลื่อนที่ของ Stepper Motor1จาก Box5_Backword" : Time;
      "เวลาเคลื่อนที่ของ Stepper Motor1จาก Box6_Backword" : Time;
      "เวลาเคลื่อนที่ของ Stepper Motor1จาก Box7_Backword" : Time;
      "เวลาเคลื่อนที่ของ Stepper Motor1จาก Box8_Backword" : Time;
      "เวลาเคลื่อนที่ของ Stepper Motor1จาก Box9_Backword" : Time;
      "เวลาเคลื่อนที่ของ Stepper Motor1จาก Box10_Backword" : Time;
      "เวลาเคลื่อนที่ของ Stepper Motor1จาก Box11_Backword" : Time;
      "เวลาเคลื่อนที่ของ Stepper Motor1จาก Box12_Backword" : Time;
      "เวลาเคลื่อนที่ของ Stepper Motor1จาก Box13_Backword" : Time;
      "เวลาเคลื่อนที่ของ Stepper Motor1จาก Box14_Backword" : Time;
      "เวลาเคลื่อนที่ของ Stepper Motor1จาก Box15_Backword" : Time;
      "เวลาเคลื่อนที่ของ Stepper Motor1จาก Box16_Backword" : Time;
      "เวลาเคลื่อนที่ของ Stepper Motor1จาก Box17_Backword" : Time;
      "เวลาเคลื่อนที่ของ Stepper Motor1จาก Box18_Backword" : Time;
      "เวลาเคลื่อนที่ของ Stepper Motor1จาก Box19_Backword" : Time;
      "เวลาเคลื่อนที่ของ Stepper Motor1จาก Box20_Backword" : Time;
   END_VAR
   VAR_IN_OUT
      "Step motor  Backword ทำงาน" : Bool;
   END_VAR
   VAR_TEMP   // added for the SCL form of the ladder/FBD networks
      _w1 : Bool;
      _w2 : Bool;
      _w3 : Bool;
      _w4 : Bool;
      _w5 : Bool;
      _w6 : Bool;
      _w7 : Bool;
      _w8 : Bool;
      _w9 : Bool;
      _w10 : Bool;
      _w11 : Bool;
      _w12 : Bool;
      _w13 : Bool;
      _w14 : Bool;
      _w15 : Bool;
      _w16 : Bool;
      _w17 : Bool;
      _w18 : Bool;
      _w19 : Bool;
      _w20 : Bool;
      _w21 : Bool;
      _w22 : Bool;
      _w23 : Bool;
      _w24 : Bool;
      _w25 : Bool;
      _w26 : Bool;
      _w27 : Bool;
      _w28 : Bool;
      _w29 : Bool;
      _w30 : Bool;
      _w31 : Bool;
      _w32 : Bool;
      _w33 : Bool;
      _w34 : Bool;
      _w35 : Bool;
      _w36 : Bool;
      _w37 : Bool;
      _w38 : Bool;
      _w39 : Bool;
   END_VAR
BEGIN

REGION Network 1
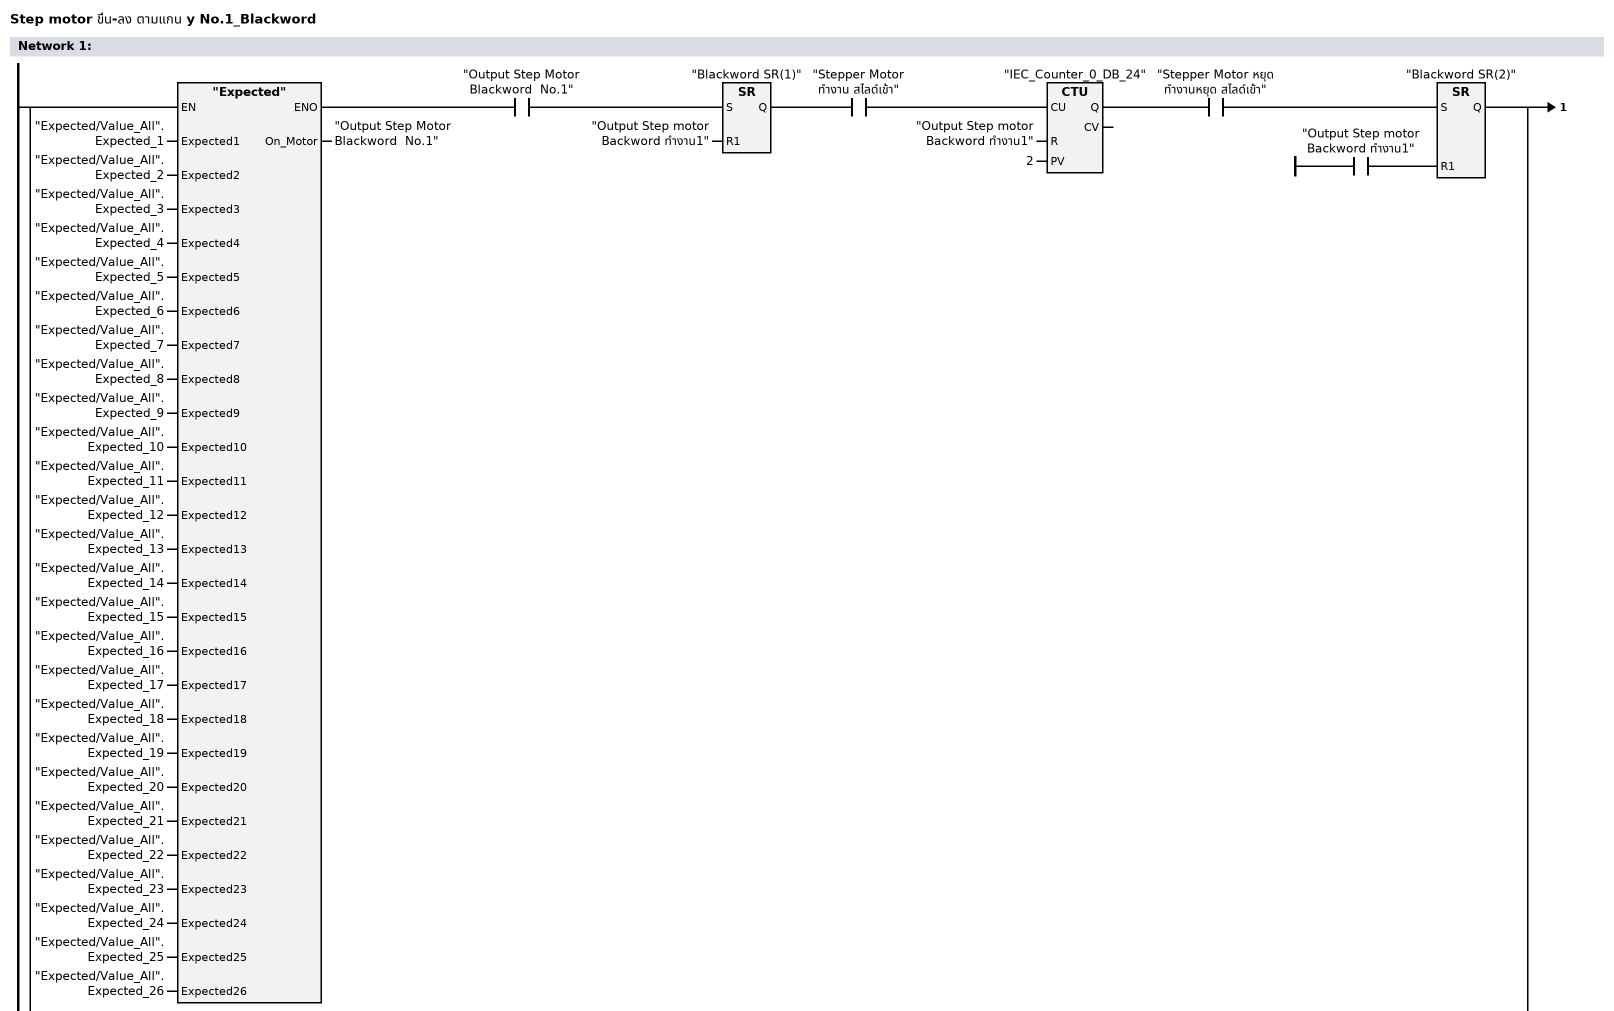
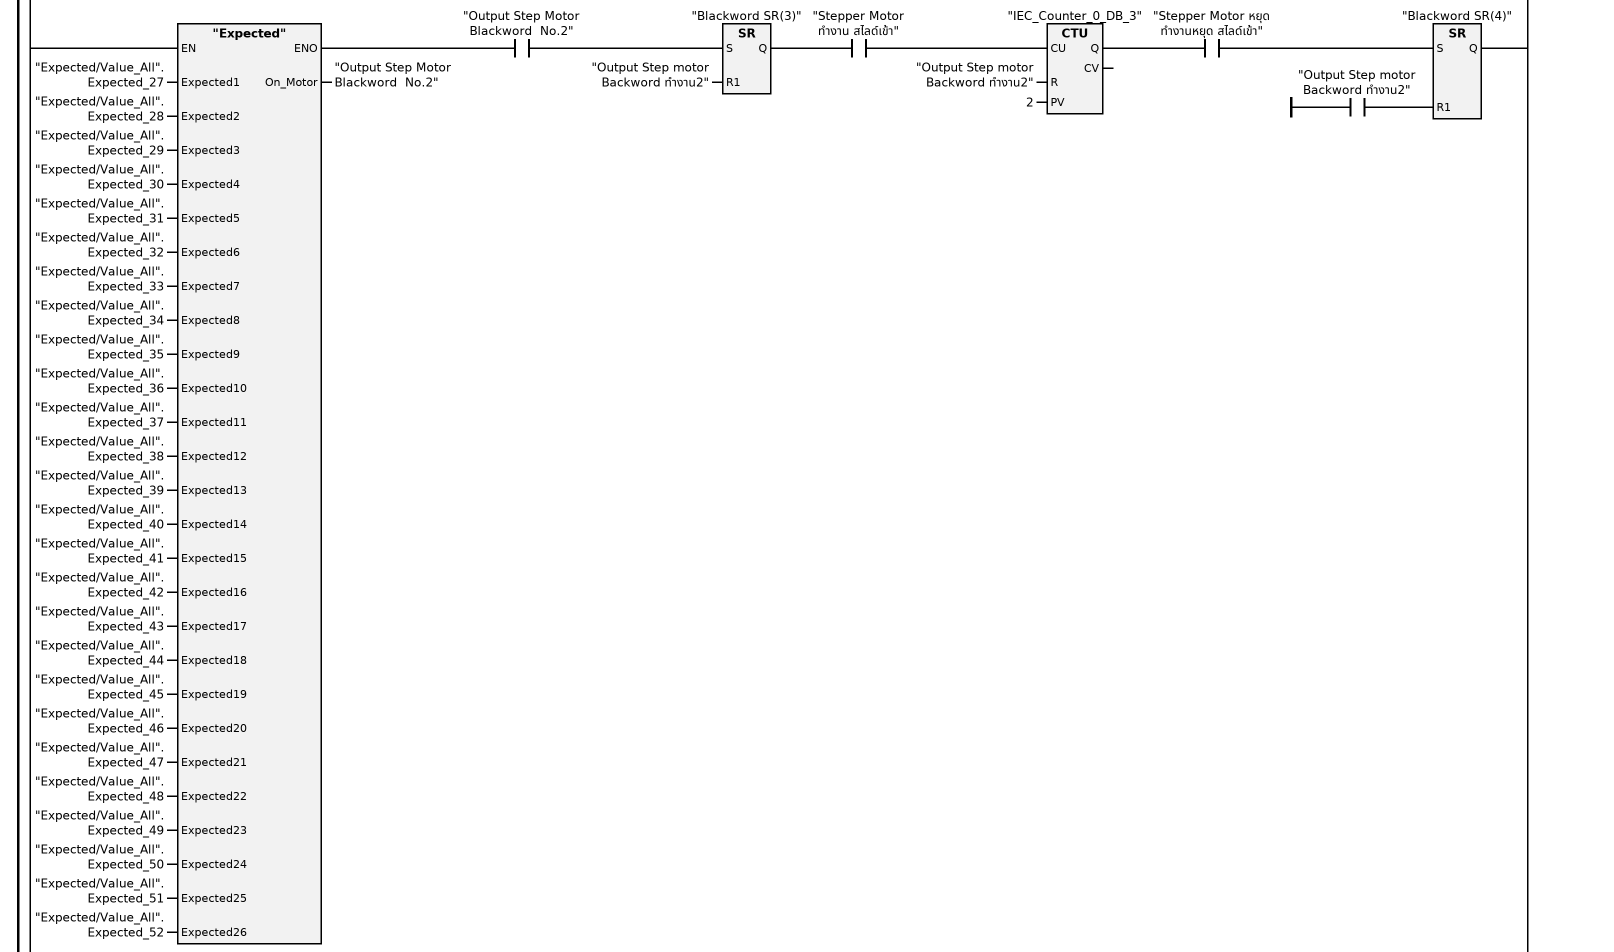
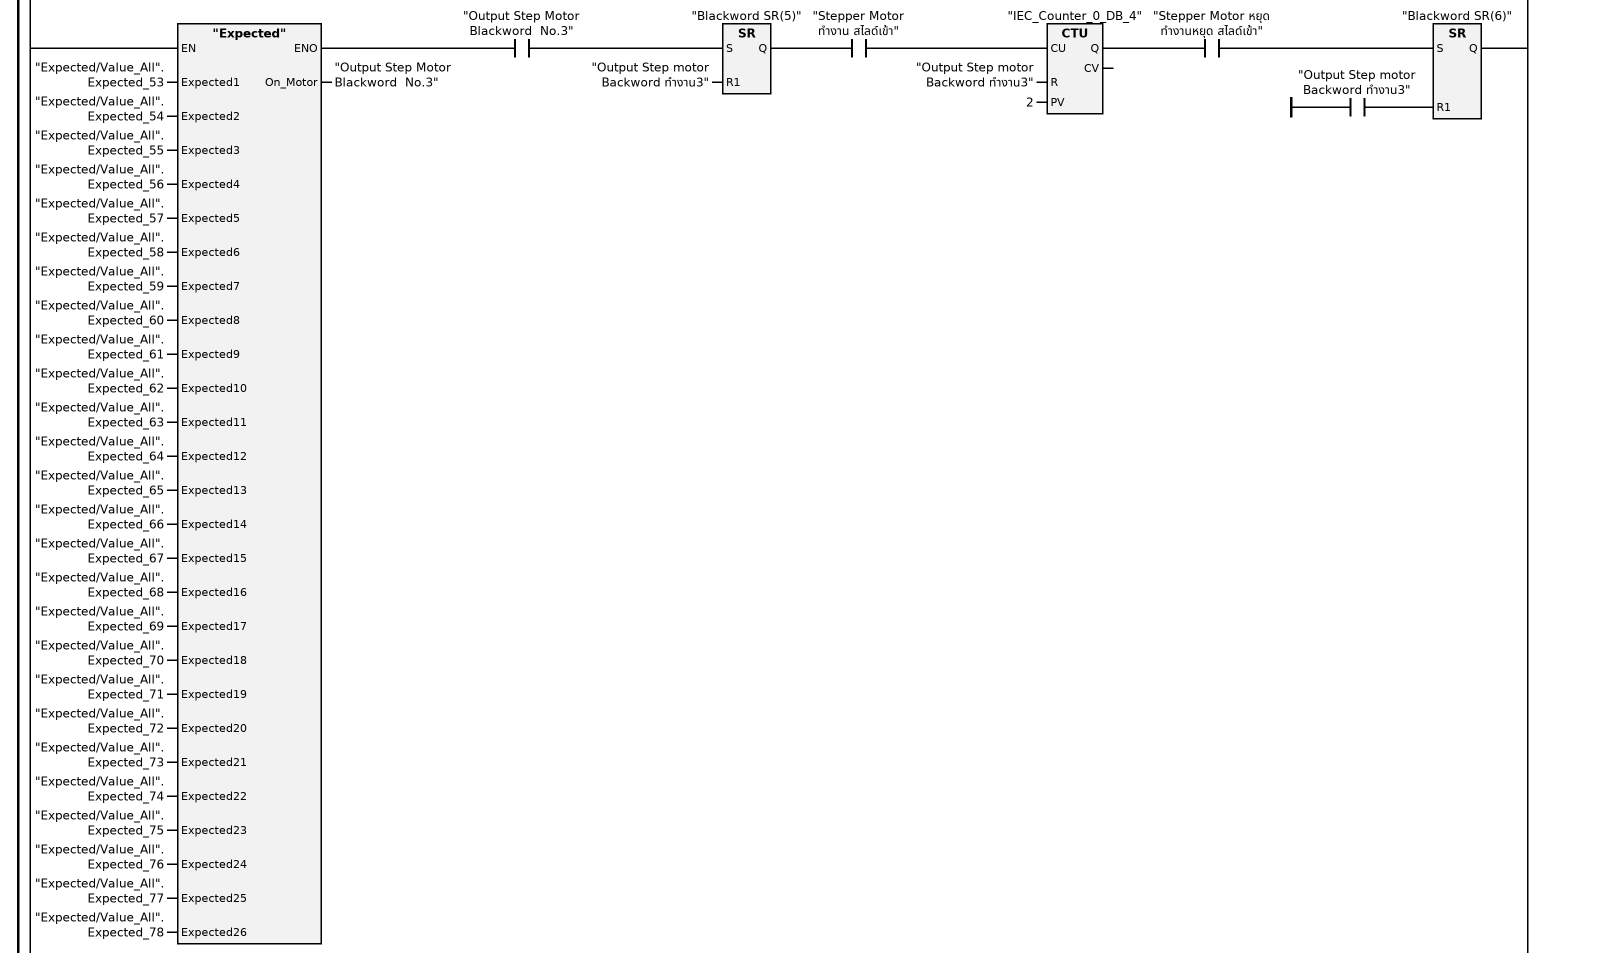
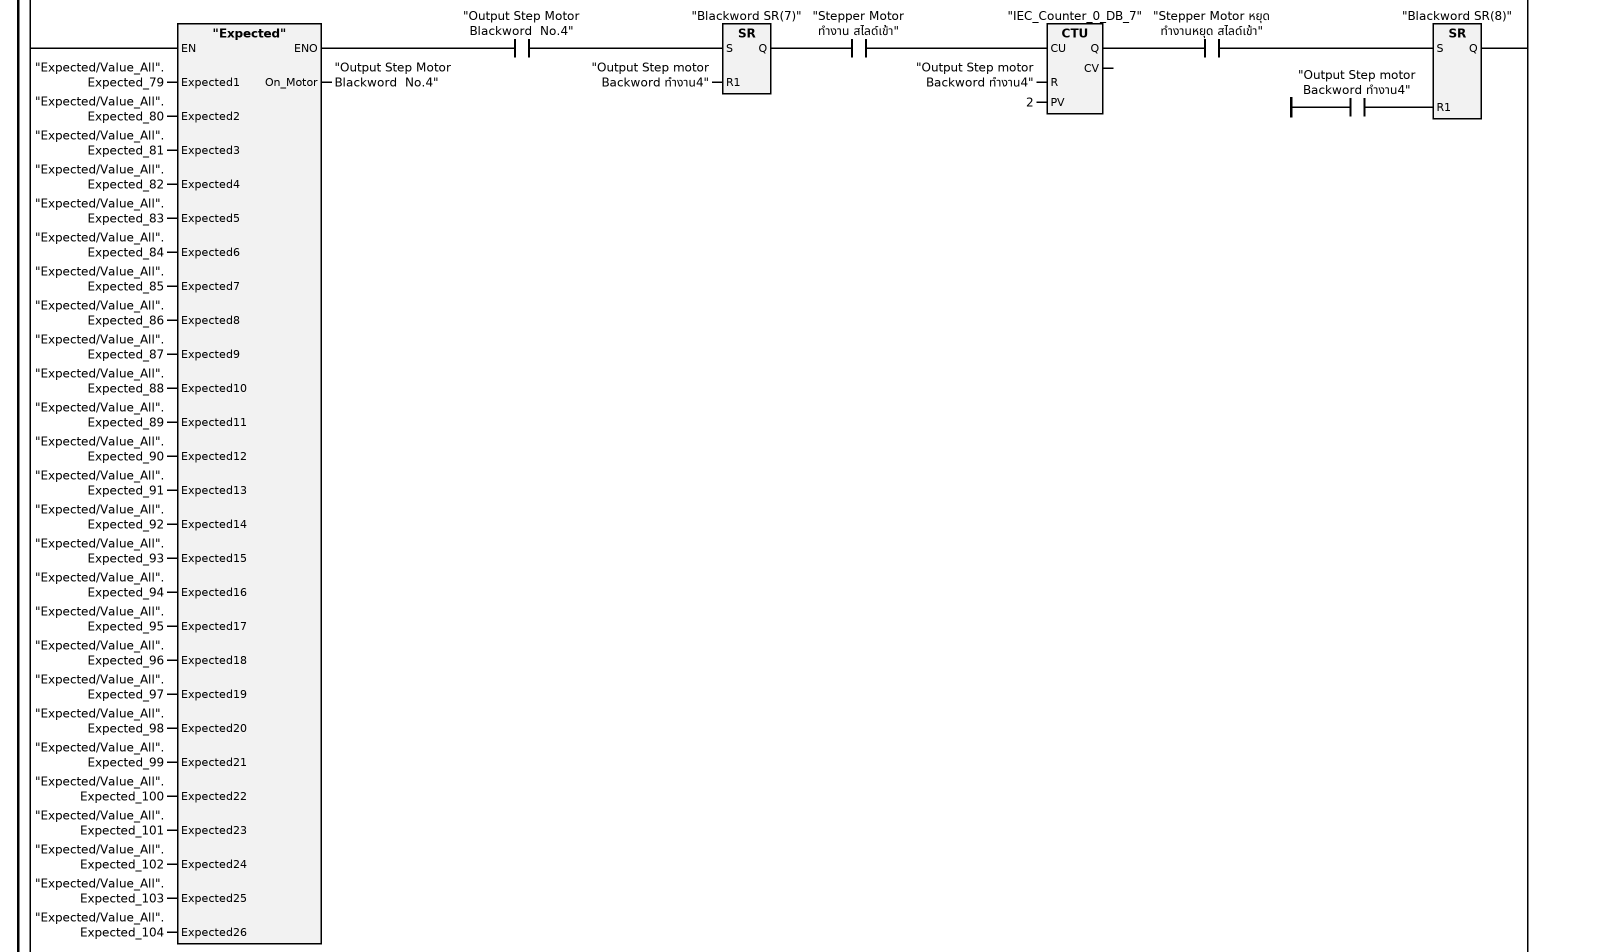
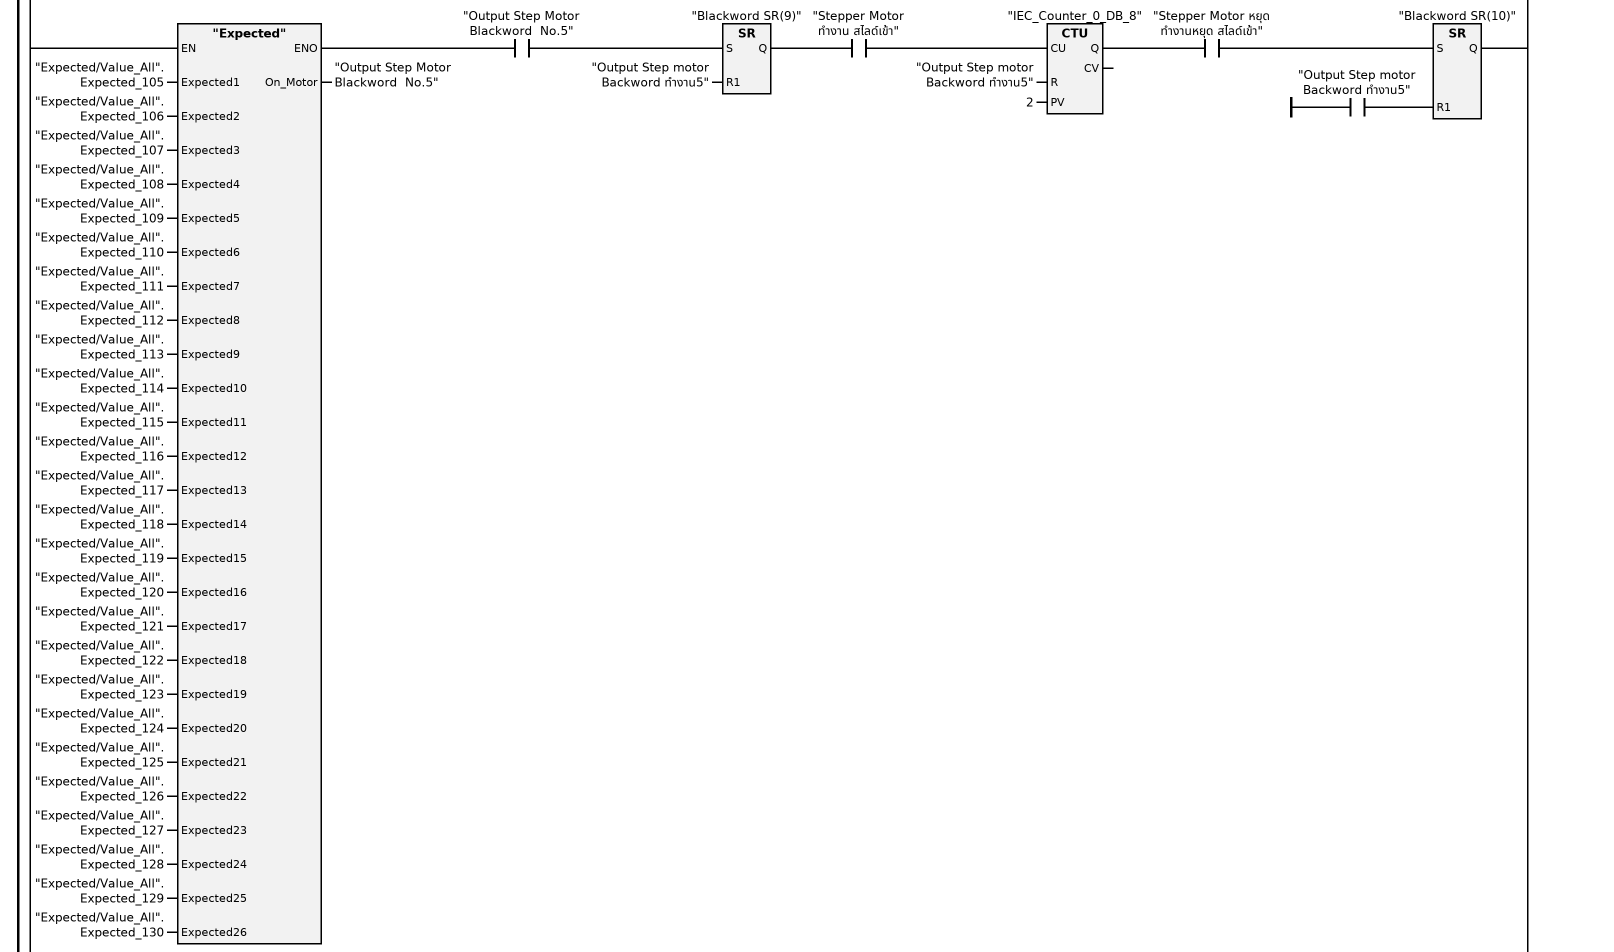
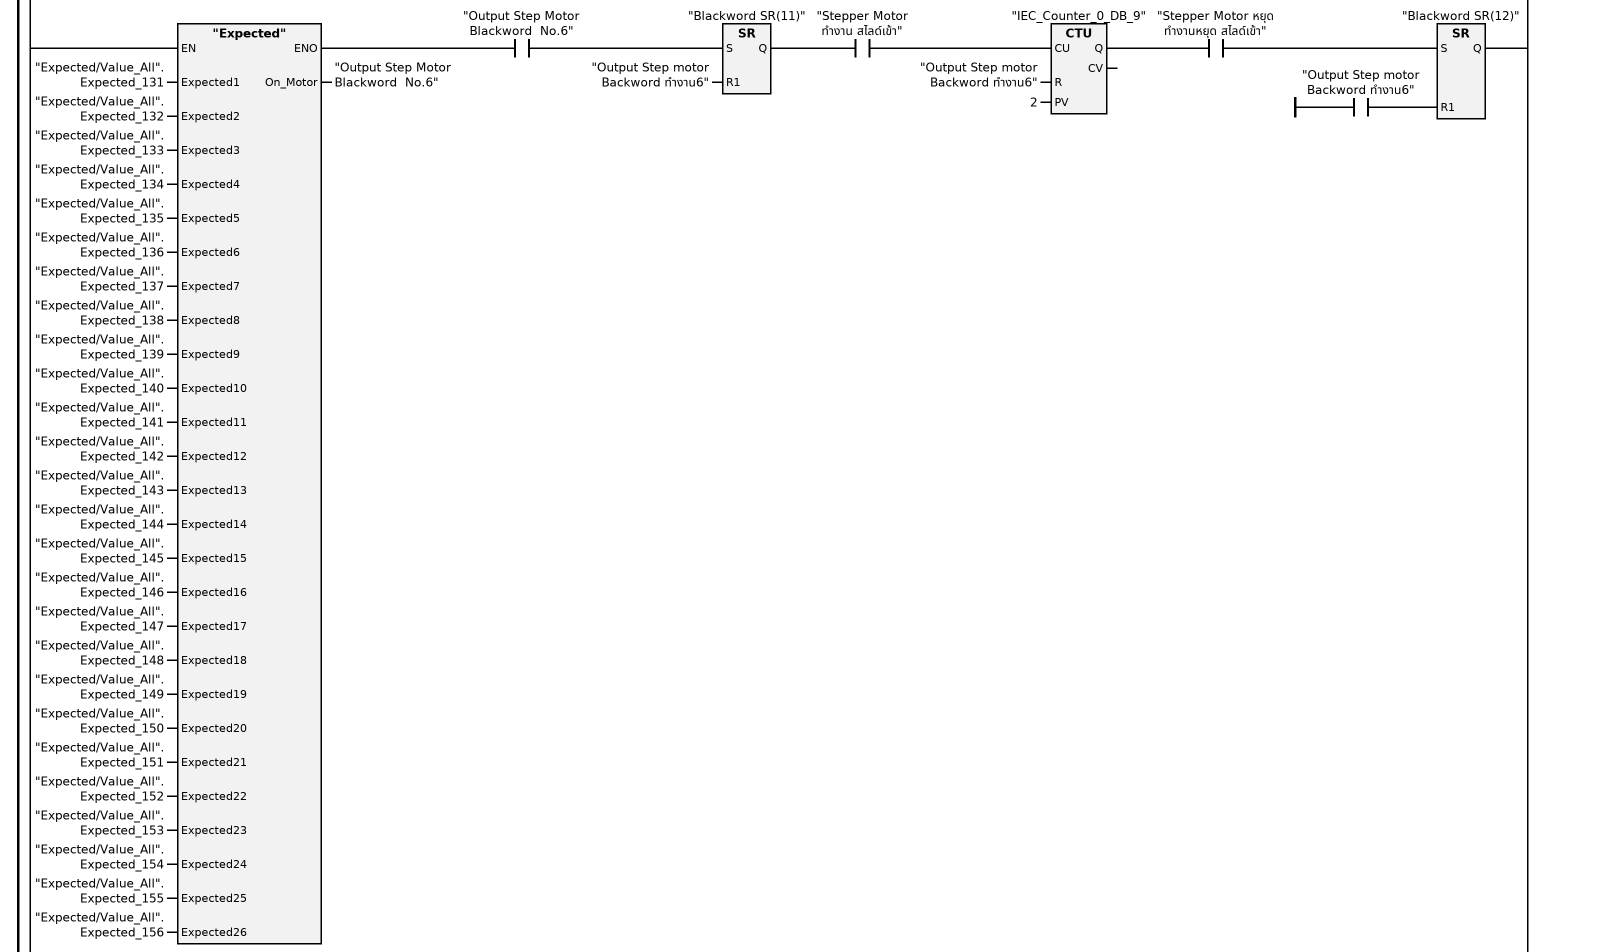
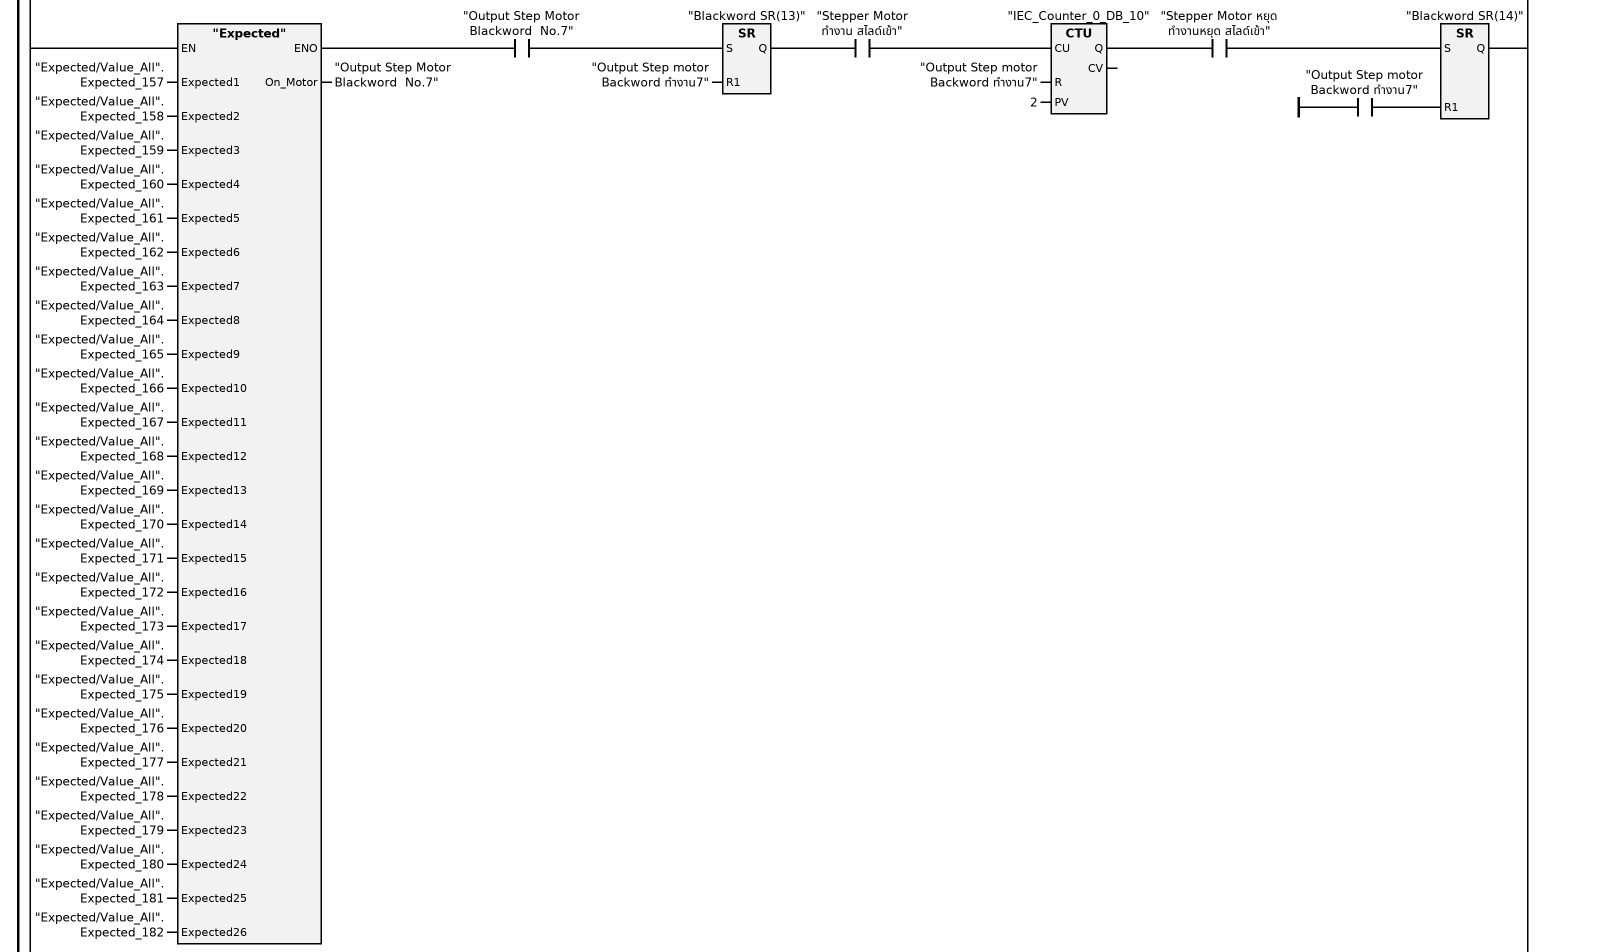
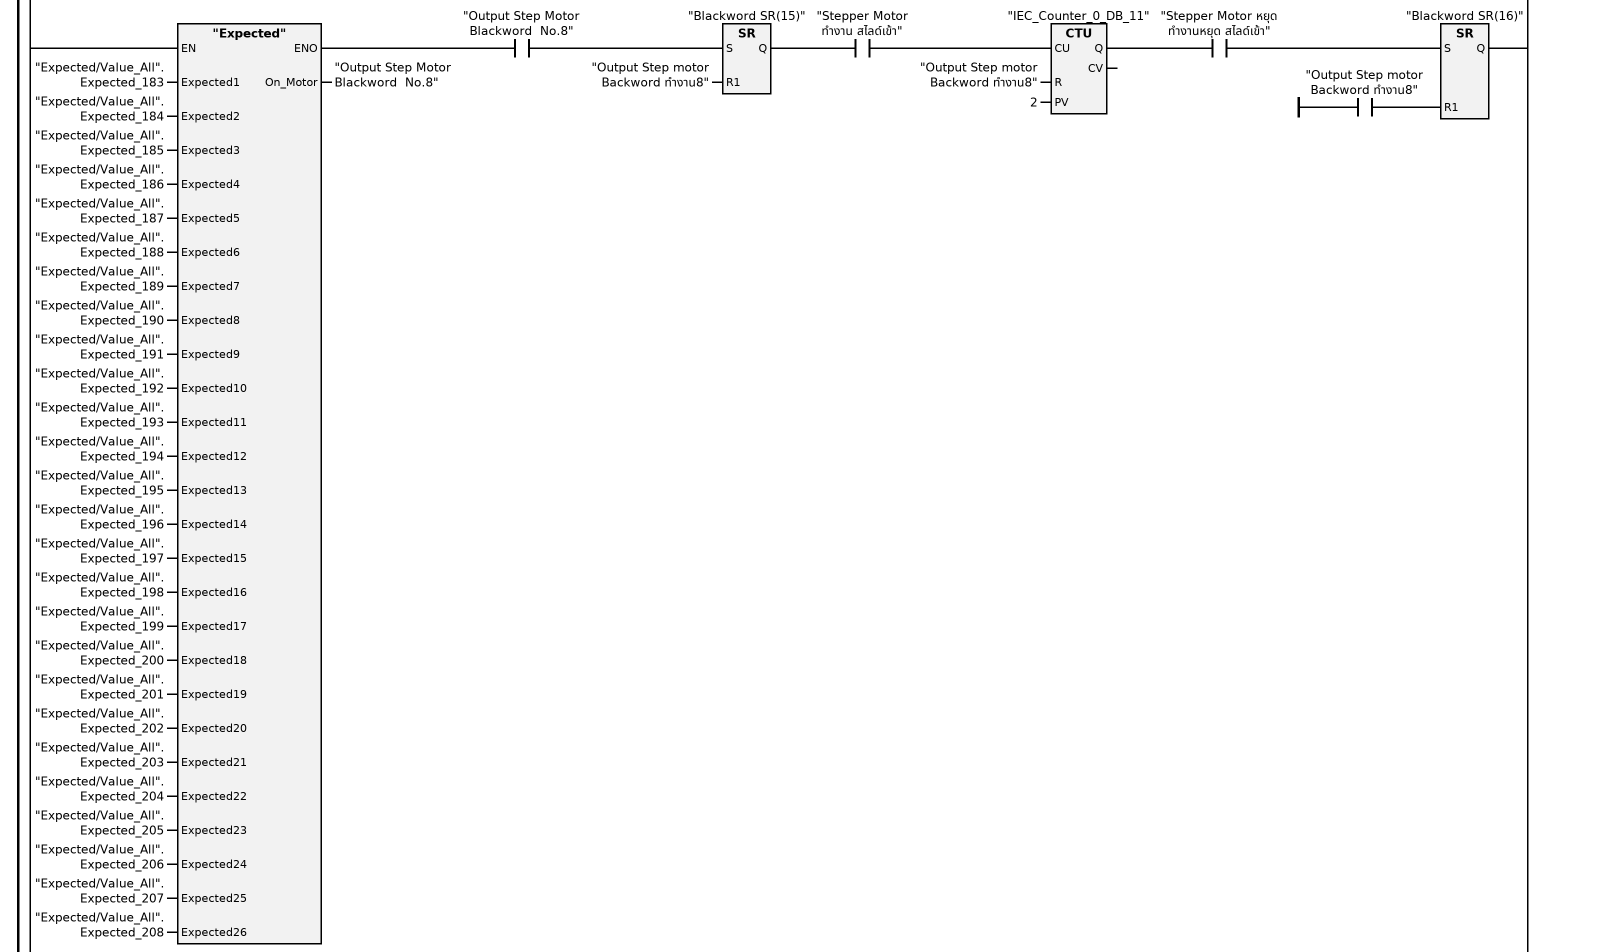
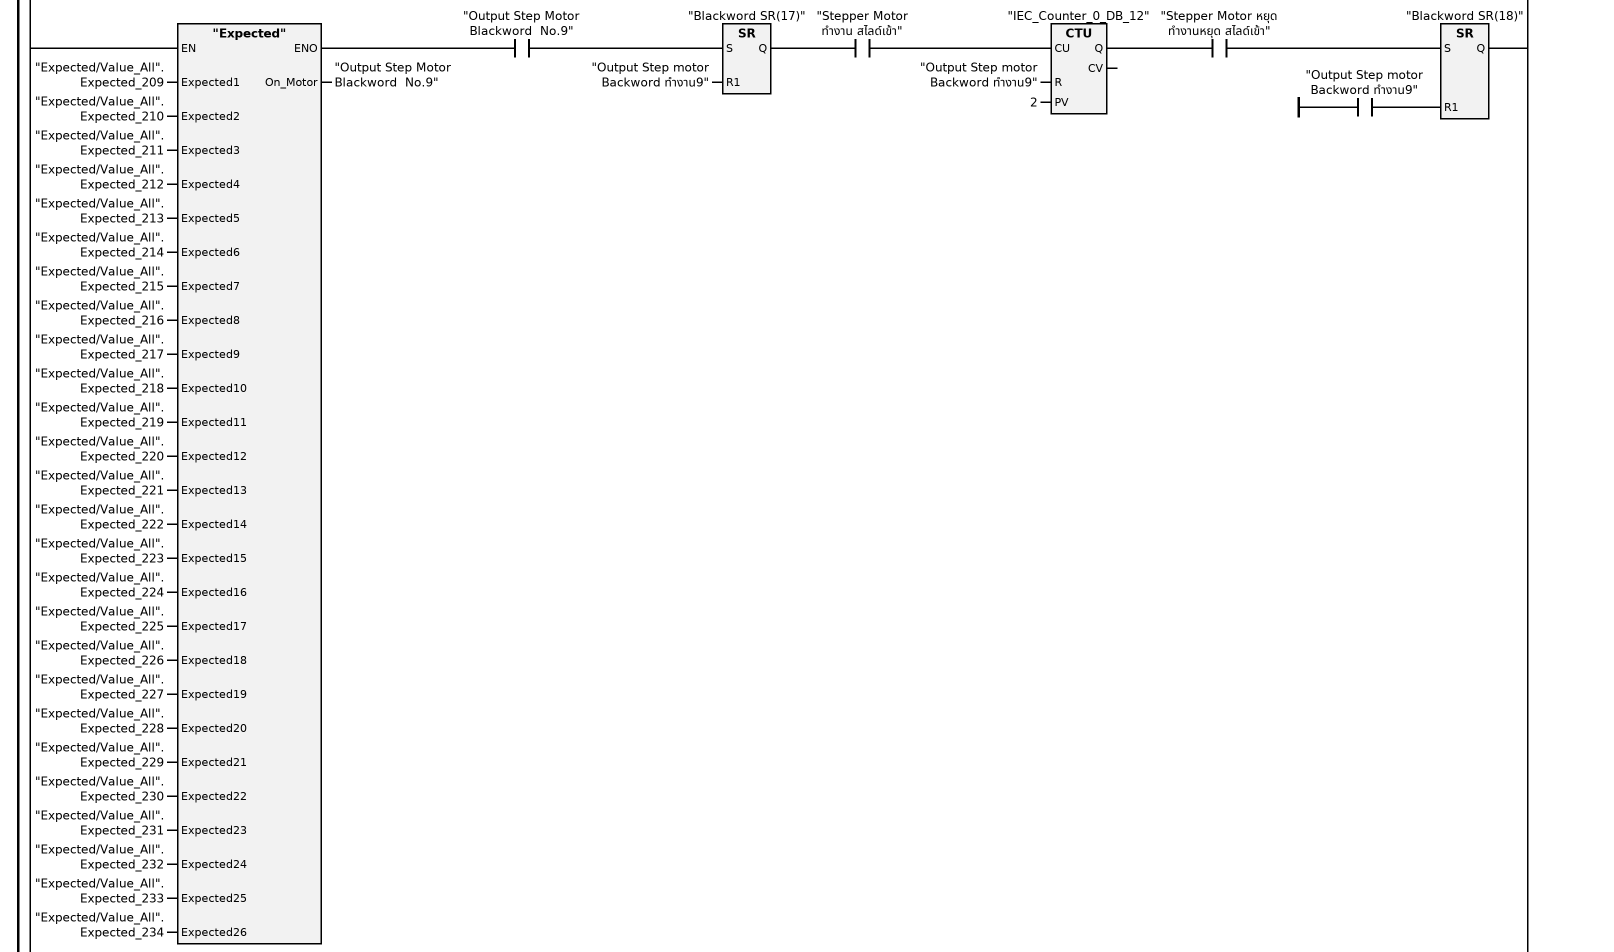
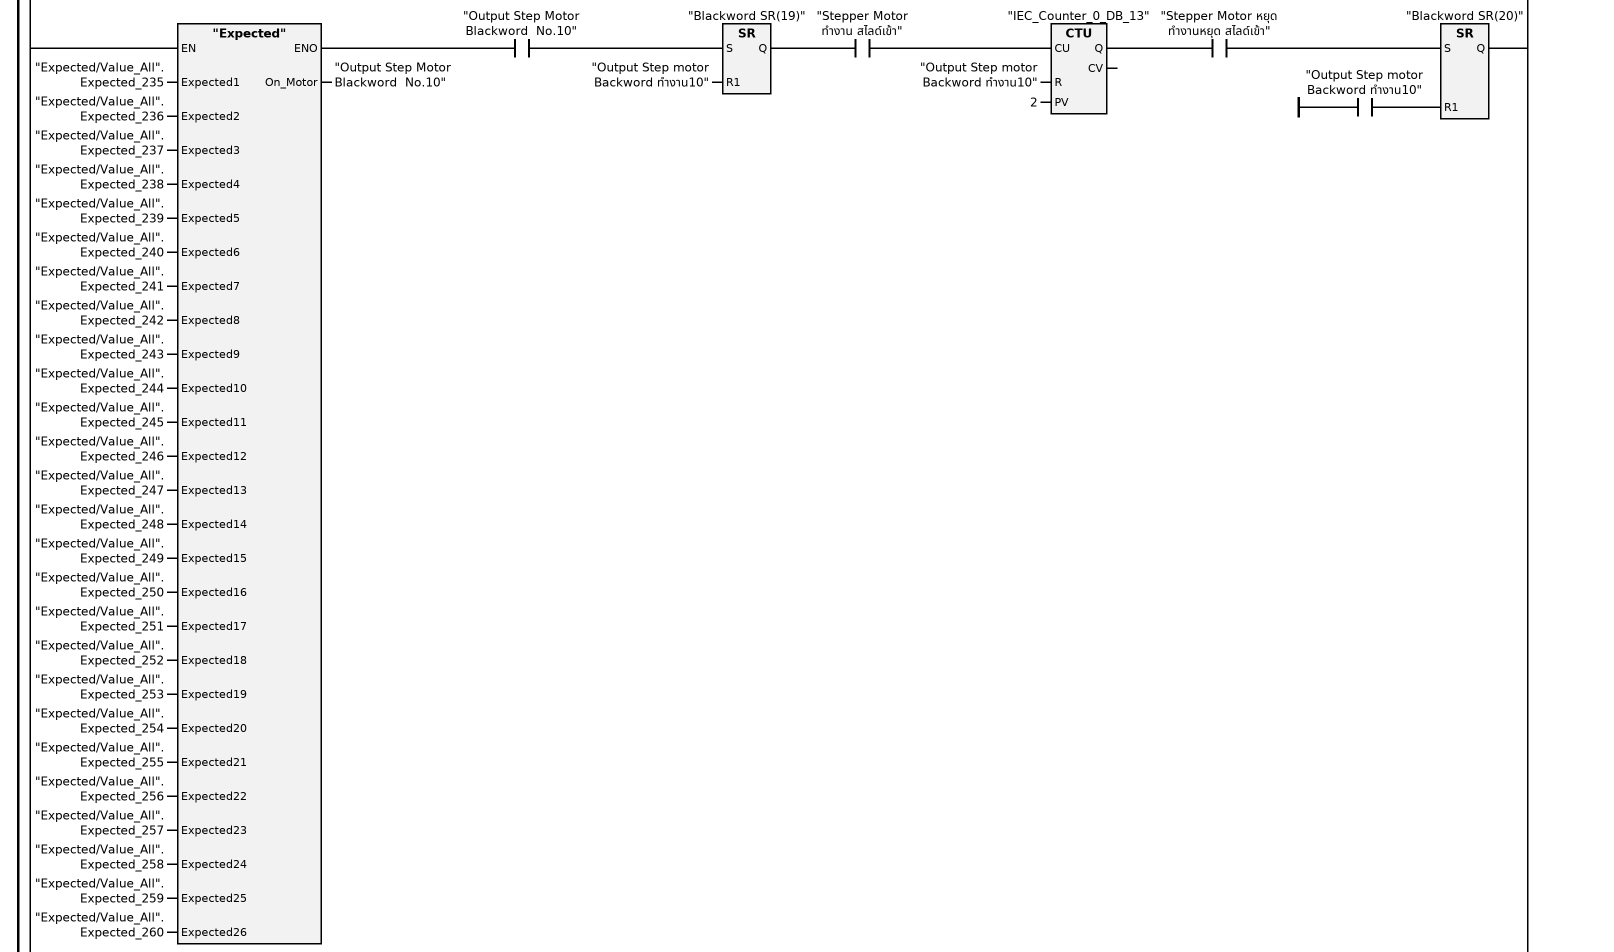
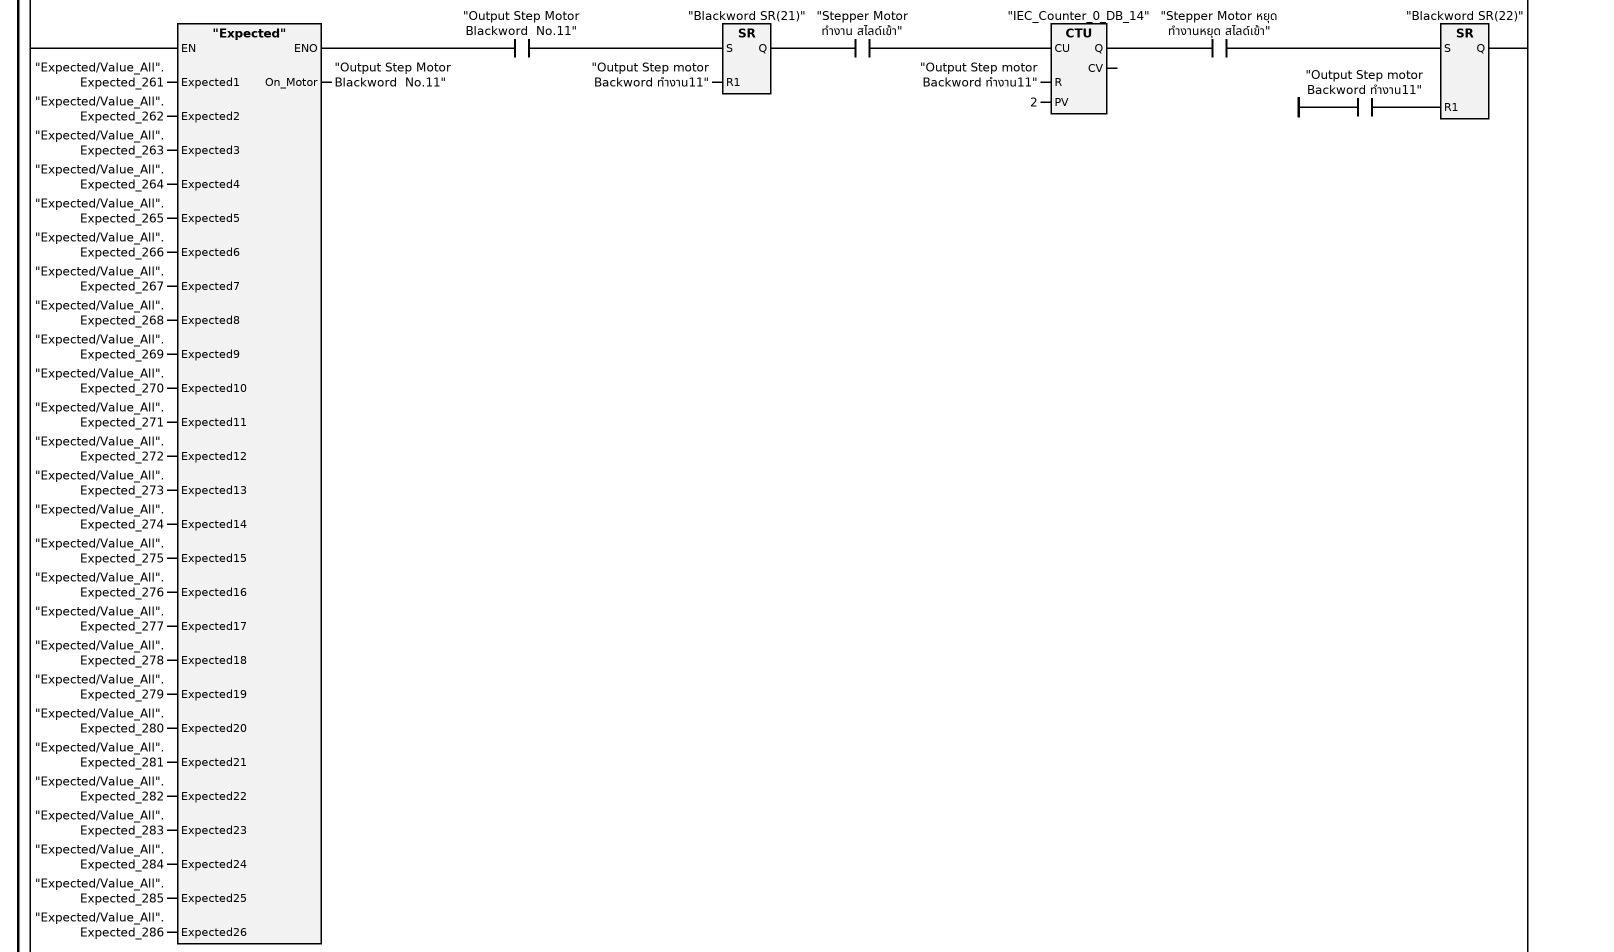
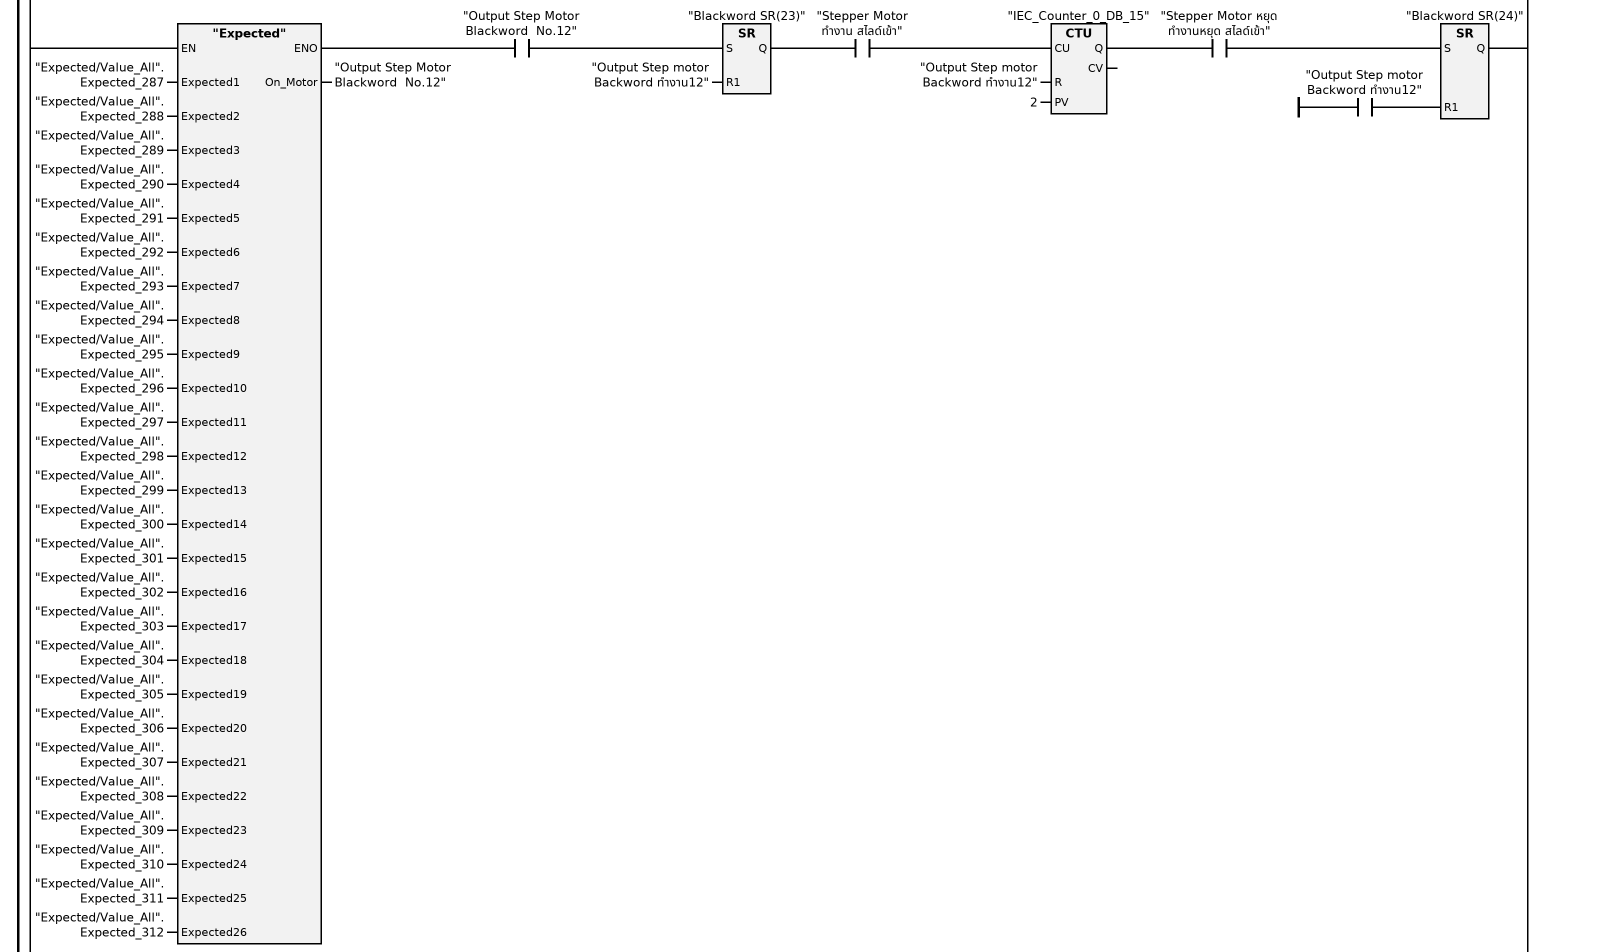
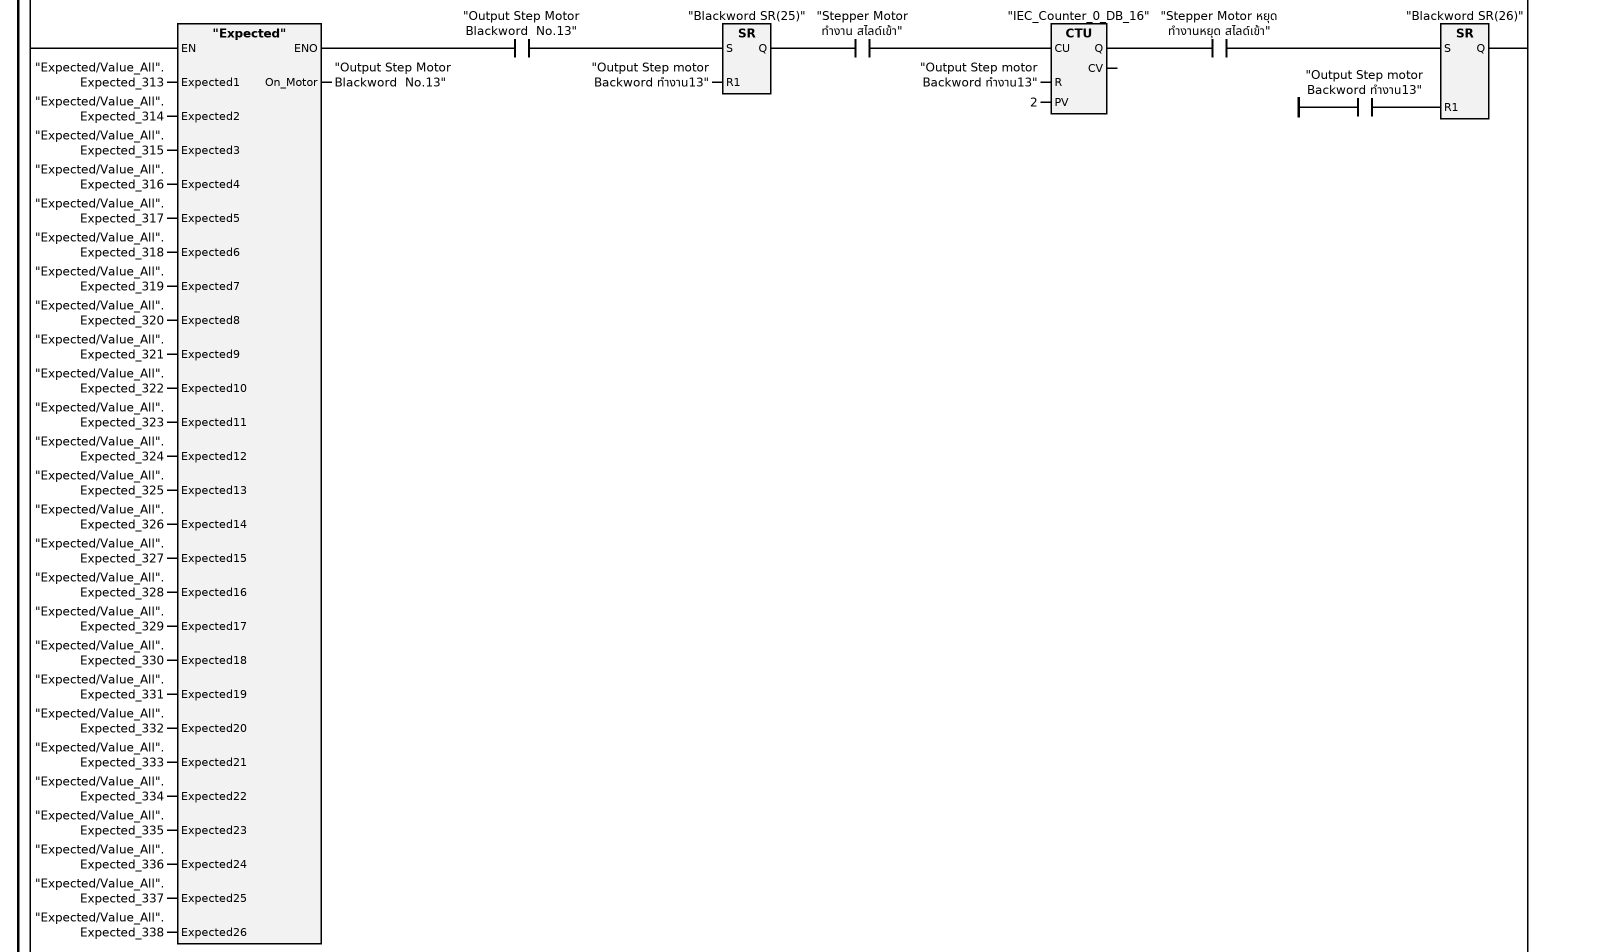
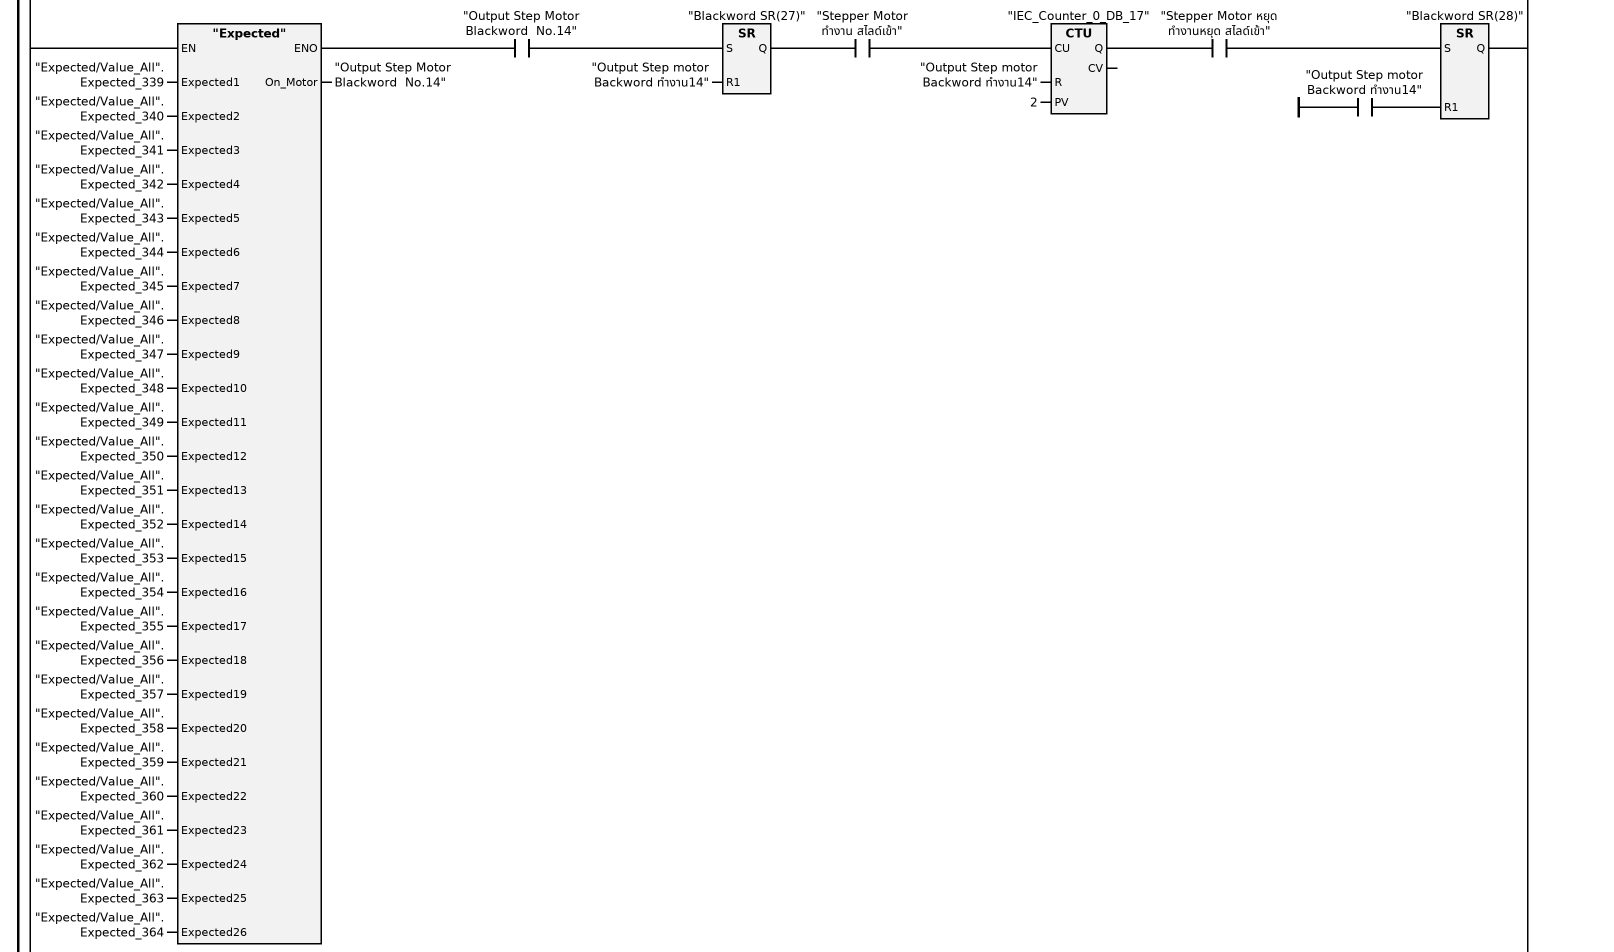
